(* CODESYS project Example15_PLC.project

Project tree, tasks and I/O mapping:
  Device : CODESYS Control Win V3, 3S - Smart Software Solutions GmbH, order no. 305021, version 3.5.7.0
    application Application
      libraries: Standard, * (System)
      task MainTask (cyclic, interval t#20ms, priority 1) calls PLC_PRG
      program PLC_PRG [ST]
      global variables GVL
      function block FB_G4LTL [ST]
    Ethernet : Ethernet, 3S - Smart Software Solutions GmbH, version 3.5.7.0
      Modbus_TCP_Master : Modbus TCP Master, 3S - Smart Software Solutions GmbH, version 3.5.6.0
          settings: AutoReconnect = TRUE
        Modbus_TCP_Slave : Modbus TCP Slave, 3S - Smart Software Solutions GmbH, version 3.5.7.0
            settings: Unit-ID = 1; IPAddress = [127, 0, 0, 1]; Channel 0.Function Code = 4; Channel 0.Read Offset = 16#0000; Channel 0.Read Length = 1; Channel 0.Write Offset = 0; Channel 0.Write Length = 0; Channel 0.Cycle Time = 100; Channel 1.Function Code = 4; Channel 1.Read Offset = 16#0001; Channel 1.Read Length = 1; Channel 1.Write Offset = 0; Channel 1.Write Length = 0; Channel 1.Cycle Time = 100; Channel 2.Function Code = 4; Channel 2.Read Offset = 16#0002; Channel 2.Read Length = 1; Channel 2.Write Offset = 0; Channel 2.Write Length = 0; Channel 2.Cycle Time = 100; Channel 3.Function Code = 4; Channel 3.Read Offset = 16#0003; Channel 3.Read Length = 1; Channel 3.Write Offset = 0; Channel 3.Write Length = 0; Channel 3.Cycle Time = 100; Channel 4.Function Code = 4; Channel 4.Read Offset = 16#0004; Channel 4.Read Length = 1; Channel 4.Write Offset = 0; Channel 4.Write Length = 0; Channel 4.Cycle Time = 100; Channel 5.Function Code = 6; Channel 5.Read Offset = 0; Channel 5.Read Length = 0; Channel 5.Write Offset = 16#0000; Channel 5.Write Length = 1; Channel 5.Cycle Time = 100; Channel 6.Function Code = 6; Channel 6.Read Offset = 0;
              Channel 6.Read Length = 0; Channel 6.Write Offset = 16#0002; Channel 6.Write Length = 1; Channel 6.Cycle Time = 100; Channel 7.Function Code = 6; Channel 7.Read Offset = 0; Channel 7.Read Length = 0; Channel 7.Write Offset = 16#0003; Channel 7.Write Length = 1; Channel 7.Cycle Time = 100; Channel 8.Function Code = 6; Channel 8.Read Offset = 0; Channel 8.Read Length = 0; Channel 8.Write Offset = 16#0004; Channel 8.Write Length = 1; Channel 8.Cycle Time = 100; Channel 9.Function Code = 6; Channel 9.Read Offset = 0; Channel 9.Read Length = 0; Channel 9.Write Offset = 16#0001; Channel 9.Write Length = 1; Channel 9.Cycle Time = 100; Channel 10.Function Code = 4; Channel 10.Read Offset = 16#0005; Channel 10.Read Length = 1; Channel 10.Write Offset = 0; Channel 10.Write Length = 0; Channel 10.Cycle Time = 100
            input  Application.dIn0 : BOOL  // Channel 0.Channel 0.Bit0
            input  Application.dIn1 : BOOL  // Channel 1.Channel 1.Bit0
            input  Application.dIn2 : BOOL  // Channel 2.Channel 2.Bit0
            input  Application.dIn3 : BOOL  // Channel 3.Channel 3.Bit0
            input  Application.dIn4 : BOOL  // Channel 4.Channel 4.Bit0
            output Application.dOut0 : BOOL  // Channel 5.Channel 5.Bit0
            output Application.dOut2 : BOOL  // Channel 6.Channel 6.Bit0
            output Application.dOut3 : BOOL  // Channel 7.Channel 7.Bit0
            output Application.dOut4 : BOOL  // Channel 8.Channel 8.Bit0
            output Application.dOut1 : BOOL  // Channel 9.Channel 9.Bit0
            input  Application.dIn5 : BOOL  // Channel 10.Channel 10.Bit0
            unmapped channels: Channel 0, Channel 1, Channel 2, Channel 3, Channel 4, Channel 5, Channel 6, Channel 7, Channel 8, Channel 9, Channel 10
*)

// Device/Application/GVL
VAR_GLOBAL
	
dIn0 : BOOL;
dIn1 : BOOL;
dIn2 : BOOL;
dIn3 : BOOL;
dIn4 : BOOL;
dIn5 : BOOL;

dOut0 : BOOL;
dOut1 : BOOL; 
dOut2 : BOOL; 
dOut3 : BOOL; 
dOut4 : BOOL; 
END_VAR

// Device/Application/PLC_PRG
PROGRAM PLC_PRG

VAR 
	fb: FB_G4LTL;
	
END_VAR


// Direct looping
// Assign pins (from global variable to function block) 
fb.x0 := dIn0;
fb.x1 := dIn1;
fb.x2 := dIn2;

// Assign pins (from function block to global variable)
dOut0 := fb.y0;
dOut1 := fb.y1;

// Run the function block
fb();

END_PROGRAM

// Device/Application/FB_G4LTL
FUNCTION_BLOCK FB_G4LTL
  (* Variable definition *)
   VAR_INPUT
      x0	: BOOL;
      x1	: BOOL;
      x2	: BOOL;
   END_VAR
   VAR_OUTPUT
      y0	: BOOL;
      y1	: BOOL;
   END_VAR
   VAR
   (* The total number of states equals to 100 *)
      cstate58	: LINT := 0;
      t0	: TON;
      t0_reset	: BOOL := FALSE;
      t0_up	: BOOL := FALSE;
      t0_start	: BOOL := FALSE;
	  
	  T0_VALUE	: TIME := TIME#7S;
   END_VAR

  (* Control logic *)
CASE cstate58 OF
1410:
    IF ((x0 = FALSE) AND  (x1 = FALSE) AND  (x2 = FALSE) AND  (t0.Q = FALSE)) THEN 
        cstate58 := 1220; y0 := FALSE; y1 := FALSE; t0_start := FALSE; 
    ELSIF ((x0 = FALSE) AND  (x1 = FALSE) AND  (x2 = FALSE) AND  (t0.Q = TRUE)) THEN 
        cstate58 := 1218; y0 := FALSE; y1 := FALSE; t0_start := FALSE; 
    ELSIF ((x0 = FALSE) AND  (x1 = FALSE) AND  (x2 = TRUE) AND  (t0.Q = FALSE)) THEN 
        cstate58 := 1412; y0 := FALSE; y1 := FALSE; t0_start := FALSE; 
    ELSIF ((x0 = FALSE) AND  (x1 = FALSE) AND  (x2 = TRUE) AND  (t0.Q = TRUE)) THEN 
        cstate58 := 1410; y0 := FALSE; y1 := FALSE; t0_start := FALSE; 
    ELSIF ((x0 = FALSE) AND  (x1 = TRUE) AND  (x2 = FALSE) AND  (t0.Q = FALSE)) THEN 
        cstate58 := 1220; y0 := FALSE; y1 := FALSE; t0_start := FALSE; 
    ELSIF ((x0 = FALSE) AND  (x1 = TRUE) AND  (x2 = FALSE) AND  (t0.Q = TRUE)) THEN 
        cstate58 := 1218; y0 := FALSE; y1 := FALSE; t0_start := FALSE; 
    ELSIF ((x0 = FALSE) AND  (x1 = TRUE) AND  (x2 = TRUE) AND  (t0.Q = FALSE)) THEN 
        cstate58 := 1412; y0 := FALSE; y1 := FALSE; t0_start := FALSE; 
    ELSIF ((x0 = FALSE) AND  (x1 = TRUE) AND  (x2 = TRUE) AND  (t0.Q = TRUE)) THEN 
        cstate58 := 1410; y0 := FALSE; y1 := FALSE; t0_start := FALSE; 
    ELSIF ((x0 = TRUE) AND  (x1 = FALSE) AND  (x2 = FALSE) AND  (t0.Q = FALSE)) THEN 
        cstate58 := 5192; y0 := TRUE; y1 := FALSE; t0_start := FALSE; 
    ELSIF ((x0 = TRUE) AND  (x1 = FALSE) AND  (x2 = FALSE) AND  (t0.Q = TRUE)) THEN 
        cstate58 := 5186; y0 := TRUE; y1 := FALSE; t0_start := FALSE; 
    ELSIF ((x0 = TRUE) AND  (x1 = FALSE) AND  (x2 = TRUE) AND  (t0.Q = FALSE)) THEN 
        cstate58 := 3848; y0 := FALSE; y1 := FALSE; t0_start := FALSE; 
    ELSIF ((x0 = TRUE) AND  (x1 = FALSE) AND  (x2 = TRUE) AND  (t0.Q = TRUE)) THEN 
        cstate58 := 3842; y0 := FALSE; y1 := FALSE; t0_start := FALSE; 
    ELSIF ((x0 = TRUE) AND  (x1 = TRUE) AND  (x2 = FALSE) AND  (t0.Q = FALSE)) THEN 
        cstate58 := 4678; y0 := TRUE; y1 := FALSE; t0_start := FALSE; 
    ELSIF ((x0 = TRUE) AND  (x1 = TRUE) AND  (x2 = FALSE) AND  (t0.Q = TRUE)) THEN 
        cstate58 := 4674; y0 := TRUE; y1 := FALSE; t0_start := FALSE; 
    ELSIF ((x0 = TRUE) AND  (x1 = TRUE) AND  (x2 = TRUE) AND  (t0.Q = FALSE)) THEN 
        cstate58 := 2502; y0 := FALSE; y1 := FALSE; t0_start := FALSE; 
    ELSIF ((x0 = TRUE) AND  (x1 = TRUE) AND  (x2 = TRUE) AND  (t0.Q = TRUE)) THEN 
        cstate58 := 2498; y0 := FALSE; y1 := FALSE; t0_start := FALSE; 
    END_IF;
6558:
    IF ((x0 = FALSE) AND  (x1 = FALSE) AND  (x2 = FALSE) AND  (t0.Q = FALSE)) THEN 
        cstate58 := 6366; y0 := FALSE; y1 := TRUE; t0_start := FALSE; 
    ELSIF ((x0 = FALSE) AND  (x1 = FALSE) AND  (x2 = FALSE) AND  (t0.Q = TRUE)) THEN 
        cstate58 := 6354; y0 := FALSE; y1 := TRUE; t0_start := FALSE; 
    ELSIF ((x0 = FALSE) AND  (x1 = FALSE) AND  (x2 = TRUE) AND  (t0.Q = FALSE)) THEN 
        cstate58 := 6558; y0 := FALSE; y1 := TRUE; t0_start := FALSE; 
    ELSIF ((x0 = FALSE) AND  (x1 = FALSE) AND  (x2 = TRUE) AND  (t0.Q = TRUE)) THEN 
        cstate58 := 6546; y0 := FALSE; y1 := TRUE; t0_start := FALSE; 
    ELSIF ((x0 = FALSE) AND  (x1 = TRUE) AND  (x2 = FALSE) AND  (t0.Q = FALSE)) THEN 
        cstate58 := 6340; y0 := FALSE; y1 := FALSE; t0_start := FALSE; 
    ELSIF ((x0 = FALSE) AND  (x1 = TRUE) AND  (x2 = FALSE) AND  (t0.Q = TRUE)) THEN 
        cstate58 := 6338; y0 := FALSE; y1 := FALSE; t0_start := FALSE; 
    ELSIF ((x0 = FALSE) AND  (x1 = TRUE) AND  (x2 = TRUE) AND  (t0.Q = FALSE)) THEN 
        cstate58 := 6532; y0 := FALSE; y1 := FALSE; t0_start := FALSE; 
    ELSIF ((x0 = FALSE) AND  (x1 = TRUE) AND  (x2 = TRUE) AND  (t0.Q = TRUE)) THEN 
        cstate58 := 6530; y0 := FALSE; y1 := FALSE; t0_start := FALSE; 
    ELSIF ((x0 = TRUE) AND  (x1 = FALSE) AND  (x2 = FALSE) AND  (t0.Q = FALSE)) THEN 
        cstate58 := 4168; y0 := TRUE; y1 := FALSE; t0_start := FALSE; 
    ELSIF ((x0 = TRUE) AND  (x1 = FALSE) AND  (x2 = FALSE) AND  (t0.Q = TRUE)) THEN 
        cstate58 := 4162; y0 := TRUE; y1 := FALSE; t0_start := FALSE; 
    ELSIF ((x0 = TRUE) AND  (x1 = FALSE) AND  (x2 = TRUE) AND  (t0.Q = FALSE)) THEN 
        cstate58 := 2824; y0 := FALSE; y1 := FALSE; t0_start := FALSE; 
    ELSIF ((x0 = TRUE) AND  (x1 = FALSE) AND  (x2 = TRUE) AND  (t0.Q = TRUE)) THEN 
        cstate58 := 2818; y0 := FALSE; y1 := FALSE; t0_start := FALSE; 
    ELSIF ((x0 = TRUE) AND  (x1 = TRUE) AND  (x2 = FALSE) AND  (t0.Q = FALSE)) THEN 
        cstate58 := 4678; y0 := TRUE; y1 := FALSE; t0_start := FALSE; 
    ELSIF ((x0 = TRUE) AND  (x1 = TRUE) AND  (x2 = FALSE) AND  (t0.Q = TRUE)) THEN 
        cstate58 := 4674; y0 := TRUE; y1 := FALSE; t0_start := FALSE; 
    ELSIF ((x0 = TRUE) AND  (x1 = TRUE) AND  (x2 = TRUE) AND  (t0.Q = FALSE)) THEN 
        cstate58 := 2502; y0 := FALSE; y1 := FALSE; t0_start := FALSE; 
    ELSIF ((x0 = TRUE) AND  (x1 = TRUE) AND  (x2 = TRUE) AND  (t0.Q = TRUE)) THEN 
        cstate58 := 2498; y0 := FALSE; y1 := FALSE; t0_start := FALSE; 
    END_IF;
1412:
    IF ((x0 = FALSE) AND  (x1 = FALSE) AND  (x2 = FALSE) AND  (t0.Q = FALSE)) THEN 
        cstate58 := 1220; y0 := FALSE; y1 := FALSE; t0_start := FALSE; 
    ELSIF ((x0 = FALSE) AND  (x1 = FALSE) AND  (x2 = FALSE) AND  (t0.Q = TRUE)) THEN 
        cstate58 := 1226; y0 := FALSE; y1 := TRUE; t0_start := FALSE; 
    ELSIF ((x0 = FALSE) AND  (x1 = FALSE) AND  (x2 = TRUE) AND  (t0.Q = FALSE)) THEN 
        cstate58 := 1412; y0 := FALSE; y1 := FALSE; t0_start := FALSE; 
    ELSIF ((x0 = FALSE) AND  (x1 = FALSE) AND  (x2 = TRUE) AND  (t0.Q = TRUE)) THEN 
        cstate58 := 1418; y0 := FALSE; y1 := TRUE; t0_start := FALSE; 
    ELSIF ((x0 = FALSE) AND  (x1 = TRUE) AND  (x2 = FALSE) AND  (t0.Q = FALSE)) THEN 
        cstate58 := 1220; y0 := FALSE; y1 := FALSE; t0_start := FALSE; 
    ELSIF ((x0 = FALSE) AND  (x1 = TRUE) AND  (x2 = FALSE) AND  (t0.Q = TRUE)) THEN 
        cstate58 := 1218; y0 := FALSE; y1 := FALSE; t0_start := FALSE; 
    ELSIF ((x0 = FALSE) AND  (x1 = TRUE) AND  (x2 = TRUE) AND  (t0.Q = FALSE)) THEN 
        cstate58 := 1412; y0 := FALSE; y1 := FALSE; t0_start := FALSE; 
    ELSIF ((x0 = FALSE) AND  (x1 = TRUE) AND  (x2 = TRUE) AND  (t0.Q = TRUE)) THEN 
        cstate58 := 1410; y0 := FALSE; y1 := FALSE; t0_start := FALSE; 
    ELSIF ((x0 = TRUE) AND  (x1 = FALSE) AND  (x2 = FALSE) AND  (t0.Q = FALSE)) THEN 
        cstate58 := 5192; y0 := TRUE; y1 := FALSE; t0_start := FALSE; 
    ELSIF ((x0 = TRUE) AND  (x1 = FALSE) AND  (x2 = FALSE) AND  (t0.Q = TRUE)) THEN 
        cstate58 := 5186; y0 := TRUE; y1 := FALSE; t0_start := FALSE; 
    ELSIF ((x0 = TRUE) AND  (x1 = FALSE) AND  (x2 = TRUE) AND  (t0.Q = FALSE)) THEN 
        cstate58 := 3848; y0 := FALSE; y1 := FALSE; t0_start := FALSE; 
    ELSIF ((x0 = TRUE) AND  (x1 = FALSE) AND  (x2 = TRUE) AND  (t0.Q = TRUE)) THEN 
        cstate58 := 3842; y0 := FALSE; y1 := FALSE; t0_start := FALSE; 
    ELSIF ((x0 = TRUE) AND  (x1 = TRUE) AND  (x2 = FALSE) AND  (t0.Q = FALSE)) THEN 
        cstate58 := 4678; y0 := TRUE; y1 := FALSE; t0_start := FALSE; 
    ELSIF ((x0 = TRUE) AND  (x1 = TRUE) AND  (x2 = FALSE) AND  (t0.Q = TRUE)) THEN 
        cstate58 := 4674; y0 := TRUE; y1 := FALSE; t0_start := FALSE; 
    ELSIF ((x0 = TRUE) AND  (x1 = TRUE) AND  (x2 = TRUE) AND  (t0.Q = FALSE)) THEN 
        cstate58 := 2502; y0 := FALSE; y1 := FALSE; t0_start := FALSE; 
    ELSIF ((x0 = TRUE) AND  (x1 = TRUE) AND  (x2 = TRUE) AND  (t0.Q = TRUE)) THEN 
        cstate58 := 2498; y0 := FALSE; y1 := FALSE; t0_start := FALSE; 
    END_IF;
1418:
    IF ((x0 = FALSE) AND  (x1 = FALSE) AND  (x2 = FALSE) AND  (t0.Q = FALSE)) THEN 
        cstate58 := 1238; y0 := FALSE; y1 := TRUE; t0_start := FALSE; 
    ELSIF ((x0 = FALSE) AND  (x1 = FALSE) AND  (x2 = FALSE) AND  (t0.Q = TRUE)) THEN 
        cstate58 := 1226; y0 := FALSE; y1 := TRUE; t0_start := FALSE; 
    ELSIF ((x0 = FALSE) AND  (x1 = FALSE) AND  (x2 = TRUE) AND  (t0.Q = FALSE)) THEN 
        cstate58 := 1430; y0 := FALSE; y1 := TRUE; t0_start := FALSE; 
    ELSIF ((x0 = FALSE) AND  (x1 = FALSE) AND  (x2 = TRUE) AND  (t0.Q = TRUE)) THEN 
        cstate58 := 1418; y0 := FALSE; y1 := TRUE; t0_start := FALSE; 
    ELSIF ((x0 = FALSE) AND  (x1 = TRUE) AND  (x2 = FALSE) AND  (t0.Q = FALSE)) THEN 
        cstate58 := 1220; y0 := FALSE; y1 := FALSE; t0_start := FALSE; 
    ELSIF ((x0 = FALSE) AND  (x1 = TRUE) AND  (x2 = FALSE) AND  (t0.Q = TRUE)) THEN 
        cstate58 := 1218; y0 := FALSE; y1 := FALSE; t0_start := FALSE; 
    ELSIF ((x0 = FALSE) AND  (x1 = TRUE) AND  (x2 = TRUE) AND  (t0.Q = FALSE)) THEN 
        cstate58 := 1412; y0 := FALSE; y1 := FALSE; t0_start := FALSE; 
    ELSIF ((x0 = FALSE) AND  (x1 = TRUE) AND  (x2 = TRUE) AND  (t0.Q = TRUE)) THEN 
        cstate58 := 1410; y0 := FALSE; y1 := FALSE; t0_start := FALSE; 
    ELSIF ((x0 = TRUE) AND  (x1 = FALSE) AND  (x2 = FALSE) AND  (t0.Q = FALSE)) THEN 
        cstate58 := 5192; y0 := TRUE; y1 := FALSE; t0_start := FALSE; 
    ELSIF ((x0 = TRUE) AND  (x1 = FALSE) AND  (x2 = FALSE) AND  (t0.Q = TRUE)) THEN 
        cstate58 := 5186; y0 := TRUE; y1 := FALSE; t0_start := FALSE; 
    ELSIF ((x0 = TRUE) AND  (x1 = FALSE) AND  (x2 = TRUE) AND  (t0.Q = FALSE)) THEN 
        cstate58 := 3848; y0 := FALSE; y1 := FALSE; t0_start := FALSE; 
    ELSIF ((x0 = TRUE) AND  (x1 = FALSE) AND  (x2 = TRUE) AND  (t0.Q = TRUE)) THEN 
        cstate58 := 3842; y0 := FALSE; y1 := FALSE; t0_start := FALSE; 
    ELSIF ((x0 = TRUE) AND  (x1 = TRUE) AND  (x2 = FALSE) AND  (t0.Q = FALSE)) THEN 
        cstate58 := 4678; y0 := TRUE; y1 := FALSE; t0_start := FALSE; 
    ELSIF ((x0 = TRUE) AND  (x1 = TRUE) AND  (x2 = FALSE) AND  (t0.Q = TRUE)) THEN 
        cstate58 := 4674; y0 := TRUE; y1 := FALSE; t0_start := FALSE; 
    ELSIF ((x0 = TRUE) AND  (x1 = TRUE) AND  (x2 = TRUE) AND  (t0.Q = FALSE)) THEN 
        cstate58 := 2502; y0 := FALSE; y1 := FALSE; t0_start := FALSE; 
    ELSIF ((x0 = TRUE) AND  (x1 = TRUE) AND  (x2 = TRUE) AND  (t0.Q = TRUE)) THEN 
        cstate58 := 2498; y0 := FALSE; y1 := FALSE; t0_start := FALSE; 
    END_IF;
7490:
    IF ((x0 = FALSE) AND  (x1 = FALSE) AND  (x2 = FALSE) AND  (t0.Q = FALSE)) THEN 
        cstate58 := 7428; y0 := FALSE; y1 := FALSE; t0_start := FALSE; 
    ELSIF ((x0 = FALSE) AND  (x1 = FALSE) AND  (x2 = FALSE) AND  (t0.Q = TRUE)) THEN 
        cstate58 := 7362; y0 := FALSE; y1 := FALSE; t0_start := FALSE; 
    ELSIF ((x0 = FALSE) AND  (x1 = FALSE) AND  (x2 = TRUE) AND  (t0.Q = FALSE)) THEN 
        cstate58 := 7492; y0 := FALSE; y1 := FALSE; t0_start := FALSE; 
    ELSIF ((x0 = FALSE) AND  (x1 = FALSE) AND  (x2 = TRUE) AND  (t0.Q = TRUE)) THEN 
        cstate58 := 7554; y0 := FALSE; y1 := FALSE; t0_start := FALSE; 
    ELSIF ((x0 = FALSE) AND  (x1 = TRUE) AND  (x2 = FALSE) AND  (t0.Q = FALSE)) THEN 
        cstate58 := 6404; y0 := FALSE; y1 := FALSE; t0_start := FALSE; 
    ELSIF ((x0 = FALSE) AND  (x1 = TRUE) AND  (x2 = FALSE) AND  (t0.Q = TRUE)) THEN 
        cstate58 := 6338; y0 := FALSE; y1 := FALSE; t0_start := FALSE; 
    ELSIF ((x0 = FALSE) AND  (x1 = TRUE) AND  (x2 = TRUE) AND  (t0.Q = FALSE)) THEN 
        cstate58 := 6468; y0 := FALSE; y1 := FALSE; t0_start := FALSE; 
    ELSIF ((x0 = FALSE) AND  (x1 = TRUE) AND  (x2 = TRUE) AND  (t0.Q = TRUE)) THEN 
        cstate58 := 6530; y0 := FALSE; y1 := FALSE; t0_start := FALSE; 
    ELSIF ((x0 = TRUE) AND  (x1 = FALSE) AND  (x2 = FALSE) AND  (t0.Q = FALSE)) THEN 
        cstate58 := 5256; y0 := TRUE; y1 := FALSE; t0_start := FALSE; 
    ELSIF ((x0 = TRUE) AND  (x1 = FALSE) AND  (x2 = FALSE) AND  (t0.Q = TRUE)) THEN 
        cstate58 := 5186; y0 := TRUE; y1 := FALSE; t0_start := FALSE; 
    ELSIF ((x0 = TRUE) AND  (x1 = FALSE) AND  (x2 = TRUE) AND  (t0.Q = FALSE)) THEN 
        cstate58 := 3784; y0 := FALSE; y1 := FALSE; t0_start := FALSE; 
    ELSIF ((x0 = TRUE) AND  (x1 = FALSE) AND  (x2 = TRUE) AND  (t0.Q = TRUE)) THEN 
        cstate58 := 3842; y0 := FALSE; y1 := FALSE; t0_start := FALSE; 
    ELSIF ((x0 = TRUE) AND  (x1 = TRUE) AND  (x2 = FALSE) AND  (t0.Q = FALSE)) THEN 
        cstate58 := 4742; y0 := TRUE; y1 := FALSE; t0_start := FALSE; 
    ELSIF ((x0 = TRUE) AND  (x1 = TRUE) AND  (x2 = FALSE) AND  (t0.Q = TRUE)) THEN 
        cstate58 := 4674; y0 := TRUE; y1 := FALSE; t0_start := FALSE; 
    ELSIF ((x0 = TRUE) AND  (x1 = TRUE) AND  (x2 = TRUE) AND  (t0.Q = FALSE)) THEN 
        cstate58 := 2566; y0 := FALSE; y1 := FALSE; t0_start := FALSE; 
    ELSIF ((x0 = TRUE) AND  (x1 = TRUE) AND  (x2 = TRUE) AND  (t0.Q = TRUE)) THEN 
        cstate58 := 2498; y0 := FALSE; y1 := FALSE; t0_start := FALSE; 
    END_IF;
7492:
    IF ((x0 = FALSE) AND  (x1 = FALSE) AND  (x2 = FALSE) AND  (t0.Q = FALSE)) THEN 
        cstate58 := 7428; y0 := FALSE; y1 := FALSE; t0_start := FALSE; 
    ELSIF ((x0 = FALSE) AND  (x1 = FALSE) AND  (x2 = FALSE) AND  (t0.Q = TRUE)) THEN 
        cstate58 := 7370; y0 := FALSE; y1 := TRUE; t0_start := FALSE; 
    ELSIF ((x0 = FALSE) AND  (x1 = FALSE) AND  (x2 = TRUE) AND  (t0.Q = FALSE)) THEN 
        cstate58 := 7492; y0 := FALSE; y1 := FALSE; t0_start := FALSE; 
    ELSIF ((x0 = FALSE) AND  (x1 = FALSE) AND  (x2 = TRUE) AND  (t0.Q = TRUE)) THEN 
        cstate58 := 7562; y0 := FALSE; y1 := TRUE; t0_start := FALSE; 
    ELSIF ((x0 = FALSE) AND  (x1 = TRUE) AND  (x2 = FALSE) AND  (t0.Q = FALSE)) THEN 
        cstate58 := 6404; y0 := FALSE; y1 := FALSE; t0_start := FALSE; 
    ELSIF ((x0 = FALSE) AND  (x1 = TRUE) AND  (x2 = FALSE) AND  (t0.Q = TRUE)) THEN 
        cstate58 := 6338; y0 := FALSE; y1 := FALSE; t0_start := FALSE; 
    ELSIF ((x0 = FALSE) AND  (x1 = TRUE) AND  (x2 = TRUE) AND  (t0.Q = FALSE)) THEN 
        cstate58 := 6468; y0 := FALSE; y1 := FALSE; t0_start := FALSE; 
    ELSIF ((x0 = FALSE) AND  (x1 = TRUE) AND  (x2 = TRUE) AND  (t0.Q = TRUE)) THEN 
        cstate58 := 6530; y0 := FALSE; y1 := FALSE; t0_start := FALSE; 
    ELSIF ((x0 = TRUE) AND  (x1 = FALSE) AND  (x2 = FALSE) AND  (t0.Q = FALSE)) THEN 
        cstate58 := 5256; y0 := TRUE; y1 := FALSE; t0_start := FALSE; 
    ELSIF ((x0 = TRUE) AND  (x1 = FALSE) AND  (x2 = FALSE) AND  (t0.Q = TRUE)) THEN 
        cstate58 := 5186; y0 := TRUE; y1 := FALSE; t0_start := FALSE; 
    ELSIF ((x0 = TRUE) AND  (x1 = FALSE) AND  (x2 = TRUE) AND  (t0.Q = FALSE)) THEN 
        cstate58 := 3784; y0 := FALSE; y1 := FALSE; t0_start := FALSE; 
    ELSIF ((x0 = TRUE) AND  (x1 = FALSE) AND  (x2 = TRUE) AND  (t0.Q = TRUE)) THEN 
        cstate58 := 3842; y0 := FALSE; y1 := FALSE; t0_start := FALSE; 
    ELSIF ((x0 = TRUE) AND  (x1 = TRUE) AND  (x2 = FALSE) AND  (t0.Q = FALSE)) THEN 
        cstate58 := 4742; y0 := TRUE; y1 := FALSE; t0_start := FALSE; 
    ELSIF ((x0 = TRUE) AND  (x1 = TRUE) AND  (x2 = FALSE) AND  (t0.Q = TRUE)) THEN 
        cstate58 := 4674; y0 := TRUE; y1 := FALSE; t0_start := FALSE; 
    ELSIF ((x0 = TRUE) AND  (x1 = TRUE) AND  (x2 = TRUE) AND  (t0.Q = FALSE)) THEN 
        cstate58 := 2566; y0 := FALSE; y1 := FALSE; t0_start := FALSE; 
    ELSIF ((x0 = TRUE) AND  (x1 = TRUE) AND  (x2 = TRUE) AND  (t0.Q = TRUE)) THEN 
        cstate58 := 2498; y0 := FALSE; y1 := FALSE; t0_start := FALSE; 
    END_IF;
6492:
    IF ((x0 = FALSE) AND  (x1 = FALSE) AND  (x2 = FALSE) AND  (t0.Q = FALSE)) THEN 
        cstate58 := 6428; y0 := FALSE; y1 := TRUE; t0_start := FALSE; 
    ELSIF ((x0 = FALSE) AND  (x1 = FALSE) AND  (x2 = FALSE) AND  (t0.Q = TRUE)) THEN 
        cstate58 := 6350; y0 := FALSE; y1 := TRUE; t0_start := FALSE; 
    ELSIF ((x0 = FALSE) AND  (x1 = FALSE) AND  (x2 = TRUE) AND  (t0.Q = FALSE)) THEN 
        cstate58 := 6492; y0 := FALSE; y1 := TRUE; t0_start := FALSE; 
    ELSIF ((x0 = FALSE) AND  (x1 = FALSE) AND  (x2 = TRUE) AND  (t0.Q = TRUE)) THEN 
        cstate58 := 6542; y0 := FALSE; y1 := TRUE; t0_start := FALSE; 
    ELSIF ((x0 = FALSE) AND  (x1 = TRUE) AND  (x2 = FALSE) AND  (t0.Q = FALSE)) THEN 
        cstate58 := 6404; y0 := FALSE; y1 := FALSE; t0_start := FALSE; 
    ELSIF ((x0 = FALSE) AND  (x1 = TRUE) AND  (x2 = FALSE) AND  (t0.Q = TRUE)) THEN 
        cstate58 := 6338; y0 := FALSE; y1 := FALSE; t0_start := FALSE; 
    ELSIF ((x0 = FALSE) AND  (x1 = TRUE) AND  (x2 = TRUE) AND  (t0.Q = FALSE)) THEN 
        cstate58 := 6468; y0 := FALSE; y1 := FALSE; t0_start := FALSE; 
    ELSIF ((x0 = FALSE) AND  (x1 = TRUE) AND  (x2 = TRUE) AND  (t0.Q = TRUE)) THEN 
        cstate58 := 6530; y0 := FALSE; y1 := FALSE; t0_start := FALSE; 
    ELSIF ((x0 = TRUE) AND  (x1 = FALSE) AND  (x2 = FALSE) AND  (t0.Q = FALSE)) THEN 
        cstate58 := 4232; y0 := TRUE; y1 := FALSE; t0_start := FALSE; 
    ELSIF ((x0 = TRUE) AND  (x1 = FALSE) AND  (x2 = FALSE) AND  (t0.Q = TRUE)) THEN 
        cstate58 := 4162; y0 := TRUE; y1 := FALSE; t0_start := FALSE; 
    ELSIF ((x0 = TRUE) AND  (x1 = FALSE) AND  (x2 = TRUE) AND  (t0.Q = FALSE)) THEN 
        cstate58 := 2760; y0 := FALSE; y1 := FALSE; t0_start := FALSE; 
    ELSIF ((x0 = TRUE) AND  (x1 = FALSE) AND  (x2 = TRUE) AND  (t0.Q = TRUE)) THEN 
        cstate58 := 2818; y0 := FALSE; y1 := FALSE; t0_start := FALSE; 
    ELSIF ((x0 = TRUE) AND  (x1 = TRUE) AND  (x2 = FALSE) AND  (t0.Q = FALSE)) THEN 
        cstate58 := 4742; y0 := TRUE; y1 := FALSE; t0_start := FALSE; 
    ELSIF ((x0 = TRUE) AND  (x1 = TRUE) AND  (x2 = FALSE) AND  (t0.Q = TRUE)) THEN 
        cstate58 := 4674; y0 := TRUE; y1 := FALSE; t0_start := FALSE; 
    ELSIF ((x0 = TRUE) AND  (x1 = TRUE) AND  (x2 = TRUE) AND  (t0.Q = FALSE)) THEN 
        cstate58 := 2566; y0 := FALSE; y1 := FALSE; t0_start := FALSE; 
    ELSIF ((x0 = TRUE) AND  (x1 = TRUE) AND  (x2 = TRUE) AND  (t0.Q = TRUE)) THEN 
        cstate58 := 2498; y0 := FALSE; y1 := FALSE; t0_start := FALSE; 
    END_IF;
6350:
    IF ((x0 = FALSE) AND  (x1 = FALSE) AND  (x2 = FALSE) AND  (t0.Q = FALSE)) THEN 
        cstate58 := 6362; y0 := FALSE; y1 := TRUE; t0_start := FALSE; 
    ELSIF ((x0 = FALSE) AND  (x1 = FALSE) AND  (x2 = FALSE) AND  (t0.Q = TRUE)) THEN 
        cstate58 := 6350; y0 := FALSE; y1 := TRUE; t0_start := FALSE; 
    ELSIF ((x0 = FALSE) AND  (x1 = FALSE) AND  (x2 = TRUE) AND  (t0.Q = FALSE)) THEN 
        cstate58 := 6492; y0 := FALSE; y1 := TRUE; t0_start := TRUE; t0_up := FALSE; 
    ELSIF ((x0 = FALSE) AND  (x1 = FALSE) AND  (x2 = TRUE) AND  (t0.Q = TRUE)) THEN 
        cstate58 := 6480; y0 := FALSE; y1 := TRUE; t0_start := TRUE; t0_up := FALSE; 
    ELSIF ((x0 = FALSE) AND  (x1 = TRUE) AND  (x2 = FALSE) AND  (t0.Q = FALSE)) THEN 
        cstate58 := 6340; y0 := FALSE; y1 := FALSE; t0_start := FALSE; 
    ELSIF ((x0 = FALSE) AND  (x1 = TRUE) AND  (x2 = FALSE) AND  (t0.Q = TRUE)) THEN 
        cstate58 := 6338; y0 := FALSE; y1 := FALSE; t0_start := FALSE; 
    ELSIF ((x0 = FALSE) AND  (x1 = TRUE) AND  (x2 = TRUE) AND  (t0.Q = FALSE)) THEN 
        cstate58 := 6468; y0 := FALSE; y1 := FALSE; t0_start := TRUE; t0_up := FALSE; 
    ELSIF ((x0 = FALSE) AND  (x1 = TRUE) AND  (x2 = TRUE) AND  (t0.Q = TRUE)) THEN 
        cstate58 := 6466; y0 := FALSE; y1 := FALSE; t0_start := TRUE; t0_up := FALSE; 
    ELSIF ((x0 = TRUE) AND  (x1 = FALSE) AND  (x2 = FALSE) AND  (t0.Q = FALSE)) THEN 
        cstate58 := 4168; y0 := TRUE; y1 := FALSE; t0_start := FALSE; 
    ELSIF ((x0 = TRUE) AND  (x1 = FALSE) AND  (x2 = FALSE) AND  (t0.Q = TRUE)) THEN 
        cstate58 := 4162; y0 := TRUE; y1 := FALSE; t0_start := FALSE; 
    ELSIF ((x0 = TRUE) AND  (x1 = FALSE) AND  (x2 = TRUE) AND  (t0.Q = FALSE)) THEN 
        cstate58 := 2760; y0 := FALSE; y1 := FALSE; t0_start := TRUE; t0_up := FALSE; 
    ELSIF ((x0 = TRUE) AND  (x1 = FALSE) AND  (x2 = TRUE) AND  (t0.Q = TRUE)) THEN 
        cstate58 := 2754; y0 := FALSE; y1 := FALSE; t0_start := TRUE; t0_up := FALSE; 
    ELSIF ((x0 = TRUE) AND  (x1 = TRUE) AND  (x2 = FALSE) AND  (t0.Q = FALSE)) THEN 
        cstate58 := 4678; y0 := TRUE; y1 := FALSE; t0_start := FALSE; 
    ELSIF ((x0 = TRUE) AND  (x1 = TRUE) AND  (x2 = FALSE) AND  (t0.Q = TRUE)) THEN 
        cstate58 := 4674; y0 := TRUE; y1 := FALSE; t0_start := FALSE; 
    ELSIF ((x0 = TRUE) AND  (x1 = TRUE) AND  (x2 = TRUE) AND  (t0.Q = FALSE)) THEN 
        cstate58 := 2566; y0 := FALSE; y1 := FALSE; t0_start := TRUE; t0_up := FALSE; 
    ELSIF ((x0 = TRUE) AND  (x1 = TRUE) AND  (x2 = TRUE) AND  (t0.Q = TRUE)) THEN 
        cstate58 := 2562; y0 := FALSE; y1 := FALSE; t0_start := TRUE; t0_up := FALSE; 
    END_IF;
6354:
    IF ((x0 = FALSE) AND  (x1 = FALSE) AND  (x2 = FALSE) AND  (t0.Q = FALSE)) THEN 
        cstate58 := 6366; y0 := FALSE; y1 := TRUE; t0_start := FALSE; 
    ELSIF ((x0 = FALSE) AND  (x1 = FALSE) AND  (x2 = FALSE) AND  (t0.Q = TRUE)) THEN 
        cstate58 := 6354; y0 := FALSE; y1 := TRUE; t0_start := FALSE; 
    ELSIF ((x0 = FALSE) AND  (x1 = FALSE) AND  (x2 = TRUE) AND  (t0.Q = FALSE)) THEN 
        cstate58 := 6496; y0 := FALSE; y1 := TRUE; t0_start := TRUE; t0_up := FALSE; 
    ELSIF ((x0 = FALSE) AND  (x1 = FALSE) AND  (x2 = TRUE) AND  (t0.Q = TRUE)) THEN 
        cstate58 := 6484; y0 := FALSE; y1 := TRUE; t0_start := TRUE; t0_up := FALSE; 
    ELSIF ((x0 = FALSE) AND  (x1 = TRUE) AND  (x2 = FALSE) AND  (t0.Q = FALSE)) THEN 
        cstate58 := 6340; y0 := FALSE; y1 := FALSE; t0_start := FALSE; 
    ELSIF ((x0 = FALSE) AND  (x1 = TRUE) AND  (x2 = FALSE) AND  (t0.Q = TRUE)) THEN 
        cstate58 := 6338; y0 := FALSE; y1 := FALSE; t0_start := FALSE; 
    ELSIF ((x0 = FALSE) AND  (x1 = TRUE) AND  (x2 = TRUE) AND  (t0.Q = FALSE)) THEN 
        cstate58 := 6468; y0 := FALSE; y1 := FALSE; t0_start := TRUE; t0_up := FALSE; 
    ELSIF ((x0 = FALSE) AND  (x1 = TRUE) AND  (x2 = TRUE) AND  (t0.Q = TRUE)) THEN 
        cstate58 := 6466; y0 := FALSE; y1 := FALSE; t0_start := TRUE; t0_up := FALSE; 
    ELSIF ((x0 = TRUE) AND  (x1 = FALSE) AND  (x2 = FALSE) AND  (t0.Q = FALSE)) THEN 
        cstate58 := 4168; y0 := TRUE; y1 := FALSE; t0_start := FALSE; 
    ELSIF ((x0 = TRUE) AND  (x1 = FALSE) AND  (x2 = FALSE) AND  (t0.Q = TRUE)) THEN 
        cstate58 := 4162; y0 := TRUE; y1 := FALSE; t0_start := FALSE; 
    ELSIF ((x0 = TRUE) AND  (x1 = FALSE) AND  (x2 = TRUE) AND  (t0.Q = FALSE)) THEN 
        cstate58 := 2760; y0 := FALSE; y1 := FALSE; t0_start := TRUE; t0_up := FALSE; 
    ELSIF ((x0 = TRUE) AND  (x1 = FALSE) AND  (x2 = TRUE) AND  (t0.Q = TRUE)) THEN 
        cstate58 := 2754; y0 := FALSE; y1 := FALSE; t0_start := TRUE; t0_up := FALSE; 
    ELSIF ((x0 = TRUE) AND  (x1 = TRUE) AND  (x2 = FALSE) AND  (t0.Q = FALSE)) THEN 
        cstate58 := 4678; y0 := TRUE; y1 := FALSE; t0_start := FALSE; 
    ELSIF ((x0 = TRUE) AND  (x1 = TRUE) AND  (x2 = FALSE) AND  (t0.Q = TRUE)) THEN 
        cstate58 := 4674; y0 := TRUE; y1 := FALSE; t0_start := FALSE; 
    ELSIF ((x0 = TRUE) AND  (x1 = TRUE) AND  (x2 = TRUE) AND  (t0.Q = FALSE)) THEN 
        cstate58 := 2566; y0 := FALSE; y1 := FALSE; t0_start := TRUE; t0_up := FALSE; 
    ELSIF ((x0 = TRUE) AND  (x1 = TRUE) AND  (x2 = TRUE) AND  (t0.Q = TRUE)) THEN 
        cstate58 := 2562; y0 := FALSE; y1 := FALSE; t0_start := TRUE; t0_up := FALSE; 
    END_IF;
6496:
    IF ((x0 = FALSE) AND  (x1 = FALSE) AND  (x2 = FALSE) AND  (t0.Q = FALSE)) THEN 
        cstate58 := 6432; y0 := FALSE; y1 := TRUE; t0_start := FALSE; 
    ELSIF ((x0 = FALSE) AND  (x1 = FALSE) AND  (x2 = FALSE) AND  (t0.Q = TRUE)) THEN 
        cstate58 := 6354; y0 := FALSE; y1 := TRUE; t0_start := FALSE; 
    ELSIF ((x0 = FALSE) AND  (x1 = FALSE) AND  (x2 = TRUE) AND  (t0.Q = FALSE)) THEN 
        cstate58 := 6496; y0 := FALSE; y1 := TRUE; t0_start := FALSE; 
    ELSIF ((x0 = FALSE) AND  (x1 = FALSE) AND  (x2 = TRUE) AND  (t0.Q = TRUE)) THEN 
        cstate58 := 6546; y0 := FALSE; y1 := TRUE; t0_start := FALSE; 
    ELSIF ((x0 = FALSE) AND  (x1 = TRUE) AND  (x2 = FALSE) AND  (t0.Q = FALSE)) THEN 
        cstate58 := 6404; y0 := FALSE; y1 := FALSE; t0_start := FALSE; 
    ELSIF ((x0 = FALSE) AND  (x1 = TRUE) AND  (x2 = FALSE) AND  (t0.Q = TRUE)) THEN 
        cstate58 := 6338; y0 := FALSE; y1 := FALSE; t0_start := FALSE; 
    ELSIF ((x0 = FALSE) AND  (x1 = TRUE) AND  (x2 = TRUE) AND  (t0.Q = FALSE)) THEN 
        cstate58 := 6468; y0 := FALSE; y1 := FALSE; t0_start := FALSE; 
    ELSIF ((x0 = FALSE) AND  (x1 = TRUE) AND  (x2 = TRUE) AND  (t0.Q = TRUE)) THEN 
        cstate58 := 6530; y0 := FALSE; y1 := FALSE; t0_start := FALSE; 
    ELSIF ((x0 = TRUE) AND  (x1 = FALSE) AND  (x2 = FALSE) AND  (t0.Q = FALSE)) THEN 
        cstate58 := 4232; y0 := TRUE; y1 := FALSE; t0_start := FALSE; 
    ELSIF ((x0 = TRUE) AND  (x1 = FALSE) AND  (x2 = FALSE) AND  (t0.Q = TRUE)) THEN 
        cstate58 := 4162; y0 := TRUE; y1 := FALSE; t0_start := FALSE; 
    ELSIF ((x0 = TRUE) AND  (x1 = FALSE) AND  (x2 = TRUE) AND  (t0.Q = FALSE)) THEN 
        cstate58 := 2760; y0 := FALSE; y1 := FALSE; t0_start := FALSE; 
    ELSIF ((x0 = TRUE) AND  (x1 = FALSE) AND  (x2 = TRUE) AND  (t0.Q = TRUE)) THEN 
        cstate58 := 2818; y0 := FALSE; y1 := FALSE; t0_start := FALSE; 
    ELSIF ((x0 = TRUE) AND  (x1 = TRUE) AND  (x2 = FALSE) AND  (t0.Q = FALSE)) THEN 
        cstate58 := 4742; y0 := TRUE; y1 := FALSE; t0_start := FALSE; 
    ELSIF ((x0 = TRUE) AND  (x1 = TRUE) AND  (x2 = FALSE) AND  (t0.Q = TRUE)) THEN 
        cstate58 := 4674; y0 := TRUE; y1 := FALSE; t0_start := FALSE; 
    ELSIF ((x0 = TRUE) AND  (x1 = TRUE) AND  (x2 = TRUE) AND  (t0.Q = FALSE)) THEN 
        cstate58 := 2566; y0 := FALSE; y1 := FALSE; t0_start := FALSE; 
    ELSIF ((x0 = TRUE) AND  (x1 = TRUE) AND  (x2 = TRUE) AND  (t0.Q = TRUE)) THEN 
        cstate58 := 2498; y0 := FALSE; y1 := FALSE; t0_start := FALSE; 
    END_IF;
6546:
    IF ((x0 = FALSE) AND  (x1 = FALSE) AND  (x2 = FALSE) AND  (t0.Q = FALSE)) THEN 
        cstate58 := 6366; y0 := FALSE; y1 := TRUE; t0_start := FALSE; 
    ELSIF ((x0 = FALSE) AND  (x1 = FALSE) AND  (x2 = FALSE) AND  (t0.Q = TRUE)) THEN 
        cstate58 := 6354; y0 := FALSE; y1 := TRUE; t0_start := FALSE; 
    ELSIF ((x0 = FALSE) AND  (x1 = FALSE) AND  (x2 = TRUE) AND  (t0.Q = FALSE)) THEN 
        cstate58 := 6558; y0 := FALSE; y1 := TRUE; t0_start := FALSE; 
    ELSIF ((x0 = FALSE) AND  (x1 = FALSE) AND  (x2 = TRUE) AND  (t0.Q = TRUE)) THEN 
        cstate58 := 6546; y0 := FALSE; y1 := TRUE; t0_start := FALSE; 
    ELSIF ((x0 = FALSE) AND  (x1 = TRUE) AND  (x2 = FALSE) AND  (t0.Q = FALSE)) THEN 
        cstate58 := 6340; y0 := FALSE; y1 := FALSE; t0_start := FALSE; 
    ELSIF ((x0 = FALSE) AND  (x1 = TRUE) AND  (x2 = FALSE) AND  (t0.Q = TRUE)) THEN 
        cstate58 := 6338; y0 := FALSE; y1 := FALSE; t0_start := FALSE; 
    ELSIF ((x0 = FALSE) AND  (x1 = TRUE) AND  (x2 = TRUE) AND  (t0.Q = FALSE)) THEN 
        cstate58 := 6532; y0 := FALSE; y1 := FALSE; t0_start := FALSE; 
    ELSIF ((x0 = FALSE) AND  (x1 = TRUE) AND  (x2 = TRUE) AND  (t0.Q = TRUE)) THEN 
        cstate58 := 6530; y0 := FALSE; y1 := FALSE; t0_start := FALSE; 
    ELSIF ((x0 = TRUE) AND  (x1 = FALSE) AND  (x2 = FALSE) AND  (t0.Q = FALSE)) THEN 
        cstate58 := 4168; y0 := TRUE; y1 := FALSE; t0_start := FALSE; 
    ELSIF ((x0 = TRUE) AND  (x1 = FALSE) AND  (x2 = FALSE) AND  (t0.Q = TRUE)) THEN 
        cstate58 := 4162; y0 := TRUE; y1 := FALSE; t0_start := FALSE; 
    ELSIF ((x0 = TRUE) AND  (x1 = FALSE) AND  (x2 = TRUE) AND  (t0.Q = FALSE)) THEN 
        cstate58 := 2824; y0 := FALSE; y1 := FALSE; t0_start := FALSE; 
    ELSIF ((x0 = TRUE) AND  (x1 = FALSE) AND  (x2 = TRUE) AND  (t0.Q = TRUE)) THEN 
        cstate58 := 2818; y0 := FALSE; y1 := FALSE; t0_start := FALSE; 
    ELSIF ((x0 = TRUE) AND  (x1 = TRUE) AND  (x2 = FALSE) AND  (t0.Q = FALSE)) THEN 
        cstate58 := 4678; y0 := TRUE; y1 := FALSE; t0_start := FALSE; 
    ELSIF ((x0 = TRUE) AND  (x1 = TRUE) AND  (x2 = FALSE) AND  (t0.Q = TRUE)) THEN 
        cstate58 := 4674; y0 := TRUE; y1 := FALSE; t0_start := FALSE; 
    ELSIF ((x0 = TRUE) AND  (x1 = TRUE) AND  (x2 = TRUE) AND  (t0.Q = FALSE)) THEN 
        cstate58 := 2502; y0 := FALSE; y1 := FALSE; t0_start := FALSE; 
    ELSIF ((x0 = TRUE) AND  (x1 = TRUE) AND  (x2 = TRUE) AND  (t0.Q = TRUE)) THEN 
        cstate58 := 2498; y0 := FALSE; y1 := FALSE; t0_start := FALSE; 
    END_IF;
1284:
    IF ((x0 = FALSE) AND  (x1 = FALSE) AND  (x2 = FALSE) AND  (t0.Q = FALSE)) THEN 
        cstate58 := 1284; y0 := FALSE; y1 := FALSE; t0_start := FALSE; 
    ELSIF ((x0 = FALSE) AND  (x1 = FALSE) AND  (x2 = FALSE) AND  (t0.Q = TRUE)) THEN 
        cstate58 := 1226; y0 := FALSE; y1 := TRUE; t0_start := FALSE; 
    ELSIF ((x0 = FALSE) AND  (x1 = FALSE) AND  (x2 = TRUE) AND  (t0.Q = FALSE)) THEN 
        cstate58 := 1348; y0 := FALSE; y1 := FALSE; t0_start := TRUE; t0_up := FALSE; 
    ELSIF ((x0 = FALSE) AND  (x1 = FALSE) AND  (x2 = TRUE) AND  (t0.Q = TRUE)) THEN 
        cstate58 := 1356; y0 := FALSE; y1 := TRUE; t0_start := TRUE; t0_up := FALSE; 
    ELSIF ((x0 = FALSE) AND  (x1 = TRUE) AND  (x2 = FALSE) AND  (t0.Q = FALSE)) THEN 
        cstate58 := 1284; y0 := FALSE; y1 := FALSE; t0_start := FALSE; 
    ELSIF ((x0 = FALSE) AND  (x1 = TRUE) AND  (x2 = FALSE) AND  (t0.Q = TRUE)) THEN 
        cstate58 := 1218; y0 := FALSE; y1 := FALSE; t0_start := FALSE; 
    ELSIF ((x0 = FALSE) AND  (x1 = TRUE) AND  (x2 = TRUE) AND  (t0.Q = FALSE)) THEN 
        cstate58 := 1348; y0 := FALSE; y1 := FALSE; t0_start := TRUE; t0_up := FALSE; 
    ELSIF ((x0 = FALSE) AND  (x1 = TRUE) AND  (x2 = TRUE) AND  (t0.Q = TRUE)) THEN 
        cstate58 := 1346; y0 := FALSE; y1 := FALSE; t0_start := TRUE; t0_up := FALSE; 
    ELSIF ((x0 = TRUE) AND  (x1 = FALSE) AND  (x2 = FALSE) AND  (t0.Q = FALSE)) THEN 
        cstate58 := 5256; y0 := TRUE; y1 := FALSE; t0_start := FALSE; 
    ELSIF ((x0 = TRUE) AND  (x1 = FALSE) AND  (x2 = FALSE) AND  (t0.Q = TRUE)) THEN 
        cstate58 := 5186; y0 := TRUE; y1 := FALSE; t0_start := FALSE; 
    ELSIF ((x0 = TRUE) AND  (x1 = FALSE) AND  (x2 = TRUE) AND  (t0.Q = FALSE)) THEN 
        cstate58 := 3784; y0 := FALSE; y1 := FALSE; t0_start := TRUE; t0_up := FALSE; 
    ELSIF ((x0 = TRUE) AND  (x1 = FALSE) AND  (x2 = TRUE) AND  (t0.Q = TRUE)) THEN 
        cstate58 := 3778; y0 := FALSE; y1 := FALSE; t0_start := TRUE; t0_up := FALSE; 
    ELSIF ((x0 = TRUE) AND  (x1 = TRUE) AND  (x2 = FALSE) AND  (t0.Q = FALSE)) THEN 
        cstate58 := 4742; y0 := TRUE; y1 := FALSE; t0_start := FALSE; 
    ELSIF ((x0 = TRUE) AND  (x1 = TRUE) AND  (x2 = FALSE) AND  (t0.Q = TRUE)) THEN 
        cstate58 := 4674; y0 := TRUE; y1 := FALSE; t0_start := FALSE; 
    ELSIF ((x0 = TRUE) AND  (x1 = TRUE) AND  (x2 = TRUE) AND  (t0.Q = FALSE)) THEN 
        cstate58 := 2566; y0 := FALSE; y1 := FALSE; t0_start := TRUE; t0_up := FALSE; 
    ELSIF ((x0 = TRUE) AND  (x1 = TRUE) AND  (x2 = TRUE) AND  (t0.Q = TRUE)) THEN 
        cstate58 := 2562; y0 := FALSE; y1 := FALSE; t0_start := TRUE; t0_up := FALSE; 
    END_IF;
3208:
    IF ((x0 = FALSE) AND  (x1 = FALSE) AND  (x2 = FALSE) AND  (t0.Q = FALSE)) THEN 
        cstate58 := 7428; y0 := FALSE; y1 := FALSE; t0_start := FALSE; 
    ELSIF ((x0 = FALSE) AND  (x1 = FALSE) AND  (x2 = FALSE) AND  (t0.Q = TRUE)) THEN 
        cstate58 := 7378; y0 := FALSE; y1 := TRUE; t0_start := FALSE; 
    ELSIF ((x0 = FALSE) AND  (x1 = FALSE) AND  (x2 = TRUE) AND  (t0.Q = FALSE)) THEN 
        cstate58 := 7492; y0 := FALSE; y1 := FALSE; t0_start := TRUE; t0_up := FALSE; 
    ELSIF ((x0 = FALSE) AND  (x1 = FALSE) AND  (x2 = TRUE) AND  (t0.Q = TRUE)) THEN 
        cstate58 := 7508; y0 := FALSE; y1 := TRUE; t0_start := TRUE; t0_up := FALSE; 
    ELSIF ((x0 = FALSE) AND  (x1 = TRUE) AND  (x2 = FALSE) AND  (t0.Q = FALSE)) THEN 
        cstate58 := 6404; y0 := FALSE; y1 := FALSE; t0_start := FALSE; 
    ELSIF ((x0 = FALSE) AND  (x1 = TRUE) AND  (x2 = FALSE) AND  (t0.Q = TRUE)) THEN 
        cstate58 := 6338; y0 := FALSE; y1 := FALSE; t0_start := FALSE; 
    ELSIF ((x0 = FALSE) AND  (x1 = TRUE) AND  (x2 = TRUE) AND  (t0.Q = FALSE)) THEN 
        cstate58 := 6468; y0 := FALSE; y1 := FALSE; t0_start := TRUE; t0_up := FALSE; 
    ELSIF ((x0 = FALSE) AND  (x1 = TRUE) AND  (x2 = TRUE) AND  (t0.Q = TRUE)) THEN 
        cstate58 := 6466; y0 := FALSE; y1 := FALSE; t0_start := TRUE; t0_up := FALSE; 
    ELSIF ((x0 = TRUE) AND  (x1 = FALSE) AND  (x2 = FALSE) AND  (t0.Q = FALSE)) THEN 
        cstate58 := 3208; y0 := FALSE; y1 := FALSE; t0_start := FALSE; 
    ELSIF ((x0 = TRUE) AND  (x1 = FALSE) AND  (x2 = FALSE) AND  (t0.Q = TRUE)) THEN 
        cstate58 := 3138; y0 := FALSE; y1 := FALSE; t0_start := FALSE; 
    ELSIF ((x0 = TRUE) AND  (x1 = FALSE) AND  (x2 = TRUE) AND  (t0.Q = FALSE)) THEN 
        cstate58 := 3784; y0 := FALSE; y1 := FALSE; t0_start := TRUE; t0_up := FALSE; 
    ELSIF ((x0 = TRUE) AND  (x1 = FALSE) AND  (x2 = TRUE) AND  (t0.Q = TRUE)) THEN 
        cstate58 := 3778; y0 := FALSE; y1 := FALSE; t0_start := TRUE; t0_up := FALSE; 
    ELSIF ((x0 = TRUE) AND  (x1 = TRUE) AND  (x2 = FALSE) AND  (t0.Q = FALSE)) THEN 
        cstate58 := 2694; y0 := FALSE; y1 := FALSE; t0_start := FALSE; 
    ELSIF ((x0 = TRUE) AND  (x1 = TRUE) AND  (x2 = FALSE) AND  (t0.Q = TRUE)) THEN 
        cstate58 := 2626; y0 := FALSE; y1 := FALSE; t0_start := FALSE; 
    ELSIF ((x0 = TRUE) AND  (x1 = TRUE) AND  (x2 = TRUE) AND  (t0.Q = FALSE)) THEN 
        cstate58 := 2566; y0 := FALSE; y1 := FALSE; t0_start := TRUE; t0_up := FALSE; 
    ELSIF ((x0 = TRUE) AND  (x1 = TRUE) AND  (x2 = TRUE) AND  (t0.Q = TRUE)) THEN 
        cstate58 := 2562; y0 := FALSE; y1 := FALSE; t0_start := TRUE; t0_up := FALSE; 
    END_IF;
3138:
    IF ((x0 = FALSE) AND  (x1 = FALSE) AND  (x2 = FALSE) AND  (t0.Q = FALSE)) THEN 
        cstate58 := 7364; y0 := FALSE; y1 := FALSE; t0_start := FALSE; 
    ELSIF ((x0 = FALSE) AND  (x1 = FALSE) AND  (x2 = FALSE) AND  (t0.Q = TRUE)) THEN 
        cstate58 := 7362; y0 := FALSE; y1 := FALSE; t0_start := FALSE; 
    ELSIF ((x0 = FALSE) AND  (x1 = FALSE) AND  (x2 = TRUE) AND  (t0.Q = FALSE)) THEN 
        cstate58 := 7492; y0 := FALSE; y1 := FALSE; t0_start := TRUE; t0_up := FALSE; 
    ELSIF ((x0 = FALSE) AND  (x1 = FALSE) AND  (x2 = TRUE) AND  (t0.Q = TRUE)) THEN 
        cstate58 := 7490; y0 := FALSE; y1 := FALSE; t0_start := TRUE; t0_up := FALSE; 
    ELSIF ((x0 = FALSE) AND  (x1 = TRUE) AND  (x2 = FALSE) AND  (t0.Q = FALSE)) THEN 
        cstate58 := 6340; y0 := FALSE; y1 := FALSE; t0_start := FALSE; 
    ELSIF ((x0 = FALSE) AND  (x1 = TRUE) AND  (x2 = FALSE) AND  (t0.Q = TRUE)) THEN 
        cstate58 := 6338; y0 := FALSE; y1 := FALSE; t0_start := FALSE; 
    ELSIF ((x0 = FALSE) AND  (x1 = TRUE) AND  (x2 = TRUE) AND  (t0.Q = FALSE)) THEN 
        cstate58 := 6468; y0 := FALSE; y1 := FALSE; t0_start := TRUE; t0_up := FALSE; 
    ELSIF ((x0 = FALSE) AND  (x1 = TRUE) AND  (x2 = TRUE) AND  (t0.Q = TRUE)) THEN 
        cstate58 := 6466; y0 := FALSE; y1 := FALSE; t0_start := TRUE; t0_up := FALSE; 
    ELSIF ((x0 = TRUE) AND  (x1 = FALSE) AND  (x2 = FALSE) AND  (t0.Q = FALSE)) THEN 
        cstate58 := 3144; y0 := FALSE; y1 := FALSE; t0_start := FALSE; 
    ELSIF ((x0 = TRUE) AND  (x1 = FALSE) AND  (x2 = FALSE) AND  (t0.Q = TRUE)) THEN 
        cstate58 := 3138; y0 := FALSE; y1 := FALSE; t0_start := FALSE; 
    ELSIF ((x0 = TRUE) AND  (x1 = FALSE) AND  (x2 = TRUE) AND  (t0.Q = FALSE)) THEN 
        cstate58 := 3784; y0 := FALSE; y1 := FALSE; t0_start := TRUE; t0_up := FALSE; 
    ELSIF ((x0 = TRUE) AND  (x1 = FALSE) AND  (x2 = TRUE) AND  (t0.Q = TRUE)) THEN 
        cstate58 := 3778; y0 := FALSE; y1 := FALSE; t0_start := TRUE; t0_up := FALSE; 
    ELSIF ((x0 = TRUE) AND  (x1 = TRUE) AND  (x2 = FALSE) AND  (t0.Q = FALSE)) THEN 
        cstate58 := 2630; y0 := FALSE; y1 := FALSE; t0_start := FALSE; 
    ELSIF ((x0 = TRUE) AND  (x1 = TRUE) AND  (x2 = FALSE) AND  (t0.Q = TRUE)) THEN 
        cstate58 := 2626; y0 := FALSE; y1 := FALSE; t0_start := FALSE; 
    ELSIF ((x0 = TRUE) AND  (x1 = TRUE) AND  (x2 = TRUE) AND  (t0.Q = FALSE)) THEN 
        cstate58 := 2566; y0 := FALSE; y1 := FALSE; t0_start := TRUE; t0_up := FALSE; 
    ELSIF ((x0 = TRUE) AND  (x1 = TRUE) AND  (x2 = TRUE) AND  (t0.Q = TRUE)) THEN 
        cstate58 := 2562; y0 := FALSE; y1 := FALSE; t0_start := TRUE; t0_up := FALSE; 
    END_IF;
6358:
    IF ((x0 = FALSE) AND  (x1 = FALSE) AND  (x2 = FALSE) AND  (t0.Q = FALSE)) THEN 
        cstate58 := 6358; y0 := FALSE; y1 := TRUE; t0_start := FALSE; 
    ELSIF ((x0 = FALSE) AND  (x1 = FALSE) AND  (x2 = FALSE) AND  (t0.Q = TRUE)) THEN 
        cstate58 := 6346; y0 := FALSE; y1 := TRUE; t0_start := FALSE; 
    ELSIF ((x0 = FALSE) AND  (x1 = FALSE) AND  (x2 = TRUE) AND  (t0.Q = FALSE)) THEN 
        cstate58 := 6488; y0 := FALSE; y1 := TRUE; t0_start := TRUE; t0_up := FALSE; 
    ELSIF ((x0 = FALSE) AND  (x1 = FALSE) AND  (x2 = TRUE) AND  (t0.Q = TRUE)) THEN 
        cstate58 := 6476; y0 := FALSE; y1 := TRUE; t0_start := TRUE; t0_up := FALSE; 
    ELSIF ((x0 = FALSE) AND  (x1 = TRUE) AND  (x2 = FALSE) AND  (t0.Q = FALSE)) THEN 
        cstate58 := 6340; y0 := FALSE; y1 := FALSE; t0_start := FALSE; 
    ELSIF ((x0 = FALSE) AND  (x1 = TRUE) AND  (x2 = FALSE) AND  (t0.Q = TRUE)) THEN 
        cstate58 := 6338; y0 := FALSE; y1 := FALSE; t0_start := FALSE; 
    ELSIF ((x0 = FALSE) AND  (x1 = TRUE) AND  (x2 = TRUE) AND  (t0.Q = FALSE)) THEN 
        cstate58 := 6468; y0 := FALSE; y1 := FALSE; t0_start := TRUE; t0_up := FALSE; 
    ELSIF ((x0 = FALSE) AND  (x1 = TRUE) AND  (x2 = TRUE) AND  (t0.Q = TRUE)) THEN 
        cstate58 := 6466; y0 := FALSE; y1 := FALSE; t0_start := TRUE; t0_up := FALSE; 
    ELSIF ((x0 = TRUE) AND  (x1 = FALSE) AND  (x2 = FALSE) AND  (t0.Q = FALSE)) THEN 
        cstate58 := 4168; y0 := TRUE; y1 := FALSE; t0_start := FALSE; 
    ELSIF ((x0 = TRUE) AND  (x1 = FALSE) AND  (x2 = FALSE) AND  (t0.Q = TRUE)) THEN 
        cstate58 := 4162; y0 := TRUE; y1 := FALSE; t0_start := FALSE; 
    ELSIF ((x0 = TRUE) AND  (x1 = FALSE) AND  (x2 = TRUE) AND  (t0.Q = FALSE)) THEN 
        cstate58 := 2760; y0 := FALSE; y1 := FALSE; t0_start := TRUE; t0_up := FALSE; 
    ELSIF ((x0 = TRUE) AND  (x1 = FALSE) AND  (x2 = TRUE) AND  (t0.Q = TRUE)) THEN 
        cstate58 := 2754; y0 := FALSE; y1 := FALSE; t0_start := TRUE; t0_up := FALSE; 
    ELSIF ((x0 = TRUE) AND  (x1 = TRUE) AND  (x2 = FALSE) AND  (t0.Q = FALSE)) THEN 
        cstate58 := 4678; y0 := TRUE; y1 := FALSE; t0_start := FALSE; 
    ELSIF ((x0 = TRUE) AND  (x1 = TRUE) AND  (x2 = FALSE) AND  (t0.Q = TRUE)) THEN 
        cstate58 := 4674; y0 := TRUE; y1 := FALSE; t0_start := FALSE; 
    ELSIF ((x0 = TRUE) AND  (x1 = TRUE) AND  (x2 = TRUE) AND  (t0.Q = FALSE)) THEN 
        cstate58 := 2566; y0 := FALSE; y1 := FALSE; t0_start := TRUE; t0_up := FALSE; 
    ELSIF ((x0 = TRUE) AND  (x1 = TRUE) AND  (x2 = TRUE) AND  (t0.Q = TRUE)) THEN 
        cstate58 := 2562; y0 := FALSE; y1 := FALSE; t0_start := TRUE; t0_up := FALSE; 
    END_IF;
2754:
    IF ((x0 = FALSE) AND  (x1 = FALSE) AND  (x2 = FALSE) AND  (t0.Q = FALSE)) THEN 
        cstate58 := 6404; y0 := FALSE; y1 := FALSE; t0_start := FALSE; 
    ELSIF ((x0 = FALSE) AND  (x1 = FALSE) AND  (x2 = FALSE) AND  (t0.Q = TRUE)) THEN 
        cstate58 := 6338; y0 := FALSE; y1 := FALSE; t0_start := FALSE; 
    ELSIF ((x0 = FALSE) AND  (x1 = FALSE) AND  (x2 = TRUE) AND  (t0.Q = FALSE)) THEN 
        cstate58 := 6468; y0 := FALSE; y1 := FALSE; t0_start := FALSE; 
    ELSIF ((x0 = FALSE) AND  (x1 = FALSE) AND  (x2 = TRUE) AND  (t0.Q = TRUE)) THEN 
        cstate58 := 6530; y0 := FALSE; y1 := FALSE; t0_start := FALSE; 
    ELSIF ((x0 = FALSE) AND  (x1 = TRUE) AND  (x2 = FALSE) AND  (t0.Q = FALSE)) THEN 
        cstate58 := 6404; y0 := FALSE; y1 := FALSE; t0_start := FALSE; 
    ELSIF ((x0 = FALSE) AND  (x1 = TRUE) AND  (x2 = FALSE) AND  (t0.Q = TRUE)) THEN 
        cstate58 := 6338; y0 := FALSE; y1 := FALSE; t0_start := FALSE; 
    ELSIF ((x0 = FALSE) AND  (x1 = TRUE) AND  (x2 = TRUE) AND  (t0.Q = FALSE)) THEN 
        cstate58 := 6468; y0 := FALSE; y1 := FALSE; t0_start := FALSE; 
    ELSIF ((x0 = FALSE) AND  (x1 = TRUE) AND  (x2 = TRUE) AND  (t0.Q = TRUE)) THEN 
        cstate58 := 6530; y0 := FALSE; y1 := FALSE; t0_start := FALSE; 
    ELSIF ((x0 = TRUE) AND  (x1 = FALSE) AND  (x2 = FALSE) AND  (t0.Q = FALSE)) THEN 
        cstate58 := 2184; y0 := FALSE; y1 := FALSE; t0_start := FALSE; 
    ELSIF ((x0 = TRUE) AND  (x1 = FALSE) AND  (x2 = FALSE) AND  (t0.Q = TRUE)) THEN 
        cstate58 := 2114; y0 := FALSE; y1 := FALSE; t0_start := FALSE; 
    ELSIF ((x0 = TRUE) AND  (x1 = FALSE) AND  (x2 = TRUE) AND  (t0.Q = FALSE)) THEN 
        cstate58 := 2760; y0 := FALSE; y1 := FALSE; t0_start := FALSE; 
    ELSIF ((x0 = TRUE) AND  (x1 = FALSE) AND  (x2 = TRUE) AND  (t0.Q = TRUE)) THEN 
        cstate58 := 2818; y0 := FALSE; y1 := FALSE; t0_start := FALSE; 
    ELSIF ((x0 = TRUE) AND  (x1 = TRUE) AND  (x2 = FALSE) AND  (t0.Q = FALSE)) THEN 
        cstate58 := 2694; y0 := FALSE; y1 := FALSE; t0_start := FALSE; 
    ELSIF ((x0 = TRUE) AND  (x1 = TRUE) AND  (x2 = FALSE) AND  (t0.Q = TRUE)) THEN 
        cstate58 := 2626; y0 := FALSE; y1 := FALSE; t0_start := FALSE; 
    ELSIF ((x0 = TRUE) AND  (x1 = TRUE) AND  (x2 = TRUE) AND  (t0.Q = FALSE)) THEN 
        cstate58 := 2566; y0 := FALSE; y1 := FALSE; t0_start := FALSE; 
    ELSIF ((x0 = TRUE) AND  (x1 = TRUE) AND  (x2 = TRUE) AND  (t0.Q = TRUE)) THEN 
        cstate58 := 2498; y0 := FALSE; y1 := FALSE; t0_start := FALSE; 
    END_IF;
6362:
    IF ((x0 = FALSE) AND  (x1 = FALSE) AND  (x2 = FALSE) AND  (t0.Q = FALSE)) THEN 
        cstate58 := 6362; y0 := FALSE; y1 := TRUE; t0_start := FALSE; 
    ELSIF ((x0 = FALSE) AND  (x1 = FALSE) AND  (x2 = FALSE) AND  (t0.Q = TRUE)) THEN 
        cstate58 := 6350; y0 := FALSE; y1 := TRUE; t0_start := FALSE; 
    ELSIF ((x0 = FALSE) AND  (x1 = FALSE) AND  (x2 = TRUE) AND  (t0.Q = FALSE)) THEN 
        cstate58 := 6492; y0 := FALSE; y1 := TRUE; t0_start := TRUE; t0_up := FALSE; 
    ELSIF ((x0 = FALSE) AND  (x1 = FALSE) AND  (x2 = TRUE) AND  (t0.Q = TRUE)) THEN 
        cstate58 := 6480; y0 := FALSE; y1 := TRUE; t0_start := TRUE; t0_up := FALSE; 
    ELSIF ((x0 = FALSE) AND  (x1 = TRUE) AND  (x2 = FALSE) AND  (t0.Q = FALSE)) THEN 
        cstate58 := 6340; y0 := FALSE; y1 := FALSE; t0_start := FALSE; 
    ELSIF ((x0 = FALSE) AND  (x1 = TRUE) AND  (x2 = FALSE) AND  (t0.Q = TRUE)) THEN 
        cstate58 := 6338; y0 := FALSE; y1 := FALSE; t0_start := FALSE; 
    ELSIF ((x0 = FALSE) AND  (x1 = TRUE) AND  (x2 = TRUE) AND  (t0.Q = FALSE)) THEN 
        cstate58 := 6468; y0 := FALSE; y1 := FALSE; t0_start := TRUE; t0_up := FALSE; 
    ELSIF ((x0 = FALSE) AND  (x1 = TRUE) AND  (x2 = TRUE) AND  (t0.Q = TRUE)) THEN 
        cstate58 := 6466; y0 := FALSE; y1 := FALSE; t0_start := TRUE; t0_up := FALSE; 
    ELSIF ((x0 = TRUE) AND  (x1 = FALSE) AND  (x2 = FALSE) AND  (t0.Q = FALSE)) THEN 
        cstate58 := 4168; y0 := TRUE; y1 := FALSE; t0_start := FALSE; 
    ELSIF ((x0 = TRUE) AND  (x1 = FALSE) AND  (x2 = FALSE) AND  (t0.Q = TRUE)) THEN 
        cstate58 := 4162; y0 := TRUE; y1 := FALSE; t0_start := FALSE; 
    ELSIF ((x0 = TRUE) AND  (x1 = FALSE) AND  (x2 = TRUE) AND  (t0.Q = FALSE)) THEN 
        cstate58 := 2760; y0 := FALSE; y1 := FALSE; t0_start := TRUE; t0_up := FALSE; 
    ELSIF ((x0 = TRUE) AND  (x1 = FALSE) AND  (x2 = TRUE) AND  (t0.Q = TRUE)) THEN 
        cstate58 := 2754; y0 := FALSE; y1 := FALSE; t0_start := TRUE; t0_up := FALSE; 
    ELSIF ((x0 = TRUE) AND  (x1 = TRUE) AND  (x2 = FALSE) AND  (t0.Q = FALSE)) THEN 
        cstate58 := 4678; y0 := TRUE; y1 := FALSE; t0_start := FALSE; 
    ELSIF ((x0 = TRUE) AND  (x1 = TRUE) AND  (x2 = FALSE) AND  (t0.Q = TRUE)) THEN 
        cstate58 := 4674; y0 := TRUE; y1 := FALSE; t0_start := FALSE; 
    ELSIF ((x0 = TRUE) AND  (x1 = TRUE) AND  (x2 = TRUE) AND  (t0.Q = FALSE)) THEN 
        cstate58 := 2566; y0 := FALSE; y1 := FALSE; t0_start := TRUE; t0_up := FALSE; 
    ELSIF ((x0 = TRUE) AND  (x1 = TRUE) AND  (x2 = TRUE) AND  (t0.Q = TRUE)) THEN 
        cstate58 := 2562; y0 := FALSE; y1 := FALSE; t0_start := TRUE; t0_up := FALSE; 
    END_IF;
6404:
    IF ((x0 = FALSE) AND  (x1 = FALSE) AND  (x2 = FALSE) AND  (t0.Q = FALSE)) THEN 
        cstate58 := 6404; y0 := FALSE; y1 := FALSE; t0_start := FALSE; 
    ELSIF ((x0 = FALSE) AND  (x1 = FALSE) AND  (x2 = FALSE) AND  (t0.Q = TRUE)) THEN 
        cstate58 := 6346; y0 := FALSE; y1 := TRUE; t0_start := FALSE; 
    ELSIF ((x0 = FALSE) AND  (x1 = FALSE) AND  (x2 = TRUE) AND  (t0.Q = FALSE)) THEN 
        cstate58 := 6468; y0 := FALSE; y1 := FALSE; t0_start := TRUE; t0_up := FALSE; 
    ELSIF ((x0 = FALSE) AND  (x1 = FALSE) AND  (x2 = TRUE) AND  (t0.Q = TRUE)) THEN 
        cstate58 := 6476; y0 := FALSE; y1 := TRUE; t0_start := TRUE; t0_up := FALSE; 
    ELSIF ((x0 = FALSE) AND  (x1 = TRUE) AND  (x2 = FALSE) AND  (t0.Q = FALSE)) THEN 
        cstate58 := 6404; y0 := FALSE; y1 := FALSE; t0_start := FALSE; 
    ELSIF ((x0 = FALSE) AND  (x1 = TRUE) AND  (x2 = FALSE) AND  (t0.Q = TRUE)) THEN 
        cstate58 := 6338; y0 := FALSE; y1 := FALSE; t0_start := FALSE; 
    ELSIF ((x0 = FALSE) AND  (x1 = TRUE) AND  (x2 = TRUE) AND  (t0.Q = FALSE)) THEN 
        cstate58 := 6468; y0 := FALSE; y1 := FALSE; t0_start := TRUE; t0_up := FALSE; 
    ELSIF ((x0 = FALSE) AND  (x1 = TRUE) AND  (x2 = TRUE) AND  (t0.Q = TRUE)) THEN 
        cstate58 := 6466; y0 := FALSE; y1 := FALSE; t0_start := TRUE; t0_up := FALSE; 
    ELSIF ((x0 = TRUE) AND  (x1 = FALSE) AND  (x2 = FALSE) AND  (t0.Q = FALSE)) THEN 
        cstate58 := 4232; y0 := TRUE; y1 := FALSE; t0_start := FALSE; 
    ELSIF ((x0 = TRUE) AND  (x1 = FALSE) AND  (x2 = FALSE) AND  (t0.Q = TRUE)) THEN 
        cstate58 := 4162; y0 := TRUE; y1 := FALSE; t0_start := FALSE; 
    ELSIF ((x0 = TRUE) AND  (x1 = FALSE) AND  (x2 = TRUE) AND  (t0.Q = FALSE)) THEN 
        cstate58 := 2760; y0 := FALSE; y1 := FALSE; t0_start := TRUE; t0_up := FALSE; 
    ELSIF ((x0 = TRUE) AND  (x1 = FALSE) AND  (x2 = TRUE) AND  (t0.Q = TRUE)) THEN 
        cstate58 := 2754; y0 := FALSE; y1 := FALSE; t0_start := TRUE; t0_up := FALSE; 
    ELSIF ((x0 = TRUE) AND  (x1 = TRUE) AND  (x2 = FALSE) AND  (t0.Q = FALSE)) THEN 
        cstate58 := 4742; y0 := TRUE; y1 := FALSE; t0_start := FALSE; 
    ELSIF ((x0 = TRUE) AND  (x1 = TRUE) AND  (x2 = FALSE) AND  (t0.Q = TRUE)) THEN 
        cstate58 := 4674; y0 := TRUE; y1 := FALSE; t0_start := FALSE; 
    ELSIF ((x0 = TRUE) AND  (x1 = TRUE) AND  (x2 = TRUE) AND  (t0.Q = FALSE)) THEN 
        cstate58 := 2566; y0 := FALSE; y1 := FALSE; t0_start := TRUE; t0_up := FALSE; 
    ELSIF ((x0 = TRUE) AND  (x1 = TRUE) AND  (x2 = TRUE) AND  (t0.Q = TRUE)) THEN 
        cstate58 := 2562; y0 := FALSE; y1 := FALSE; t0_start := TRUE; t0_up := FALSE; 
    END_IF;
0:
    IF ((x0 = FALSE) AND  (x1 = FALSE) AND  (x2 = FALSE) AND  (t0.Q = FALSE)) THEN 
        cstate58 := 1220; y0 := FALSE; y1 := FALSE; t0_start := FALSE; 
    ELSIF ((x0 = FALSE) AND  (x1 = FALSE) AND  (x2 = FALSE) AND  (t0.Q = TRUE)) THEN 
        cstate58 := 1218; y0 := FALSE; y1 := FALSE; t0_start := FALSE; 
    ELSIF ((x0 = FALSE) AND  (x1 = FALSE) AND  (x2 = TRUE) AND  (t0.Q = FALSE)) THEN 
        cstate58 := 1412; y0 := FALSE; y1 := FALSE; t0_start := FALSE; 
    ELSIF ((x0 = FALSE) AND  (x1 = FALSE) AND  (x2 = TRUE) AND  (t0.Q = TRUE)) THEN 
        cstate58 := 1410; y0 := FALSE; y1 := FALSE; t0_start := FALSE; 
    ELSIF ((x0 = FALSE) AND  (x1 = TRUE) AND  (x2 = FALSE) AND  (t0.Q = FALSE)) THEN 
        cstate58 := 1220; y0 := FALSE; y1 := FALSE; t0_start := FALSE; 
    ELSIF ((x0 = FALSE) AND  (x1 = TRUE) AND  (x2 = FALSE) AND  (t0.Q = TRUE)) THEN 
        cstate58 := 1218; y0 := FALSE; y1 := FALSE; t0_start := FALSE; 
    ELSIF ((x0 = FALSE) AND  (x1 = TRUE) AND  (x2 = TRUE) AND  (t0.Q = FALSE)) THEN 
        cstate58 := 1412; y0 := FALSE; y1 := FALSE; t0_start := FALSE; 
    ELSIF ((x0 = FALSE) AND  (x1 = TRUE) AND  (x2 = TRUE) AND  (t0.Q = TRUE)) THEN 
        cstate58 := 1410; y0 := FALSE; y1 := FALSE; t0_start := FALSE; 
    ELSIF ((x0 = TRUE) AND  (x1 = FALSE) AND  (x2 = FALSE) AND  (t0.Q = FALSE)) THEN 
        cstate58 := 3144; y0 := FALSE; y1 := FALSE; t0_start := FALSE; 
    ELSIF ((x0 = TRUE) AND  (x1 = FALSE) AND  (x2 = FALSE) AND  (t0.Q = TRUE)) THEN 
        cstate58 := 3138; y0 := FALSE; y1 := FALSE; t0_start := FALSE; 
    ELSIF ((x0 = TRUE) AND  (x1 = FALSE) AND  (x2 = TRUE) AND  (t0.Q = FALSE)) THEN 
        cstate58 := 3848; y0 := FALSE; y1 := FALSE; t0_start := FALSE; 
    ELSIF ((x0 = TRUE) AND  (x1 = FALSE) AND  (x2 = TRUE) AND  (t0.Q = TRUE)) THEN 
        cstate58 := 3842; y0 := FALSE; y1 := FALSE; t0_start := FALSE; 
    ELSIF ((x0 = TRUE) AND  (x1 = TRUE) AND  (x2 = FALSE) AND  (t0.Q = FALSE)) THEN 
        cstate58 := 2630; y0 := FALSE; y1 := FALSE; t0_start := FALSE; 
    ELSIF ((x0 = TRUE) AND  (x1 = TRUE) AND  (x2 = FALSE) AND  (t0.Q = TRUE)) THEN 
        cstate58 := 2626; y0 := FALSE; y1 := FALSE; t0_start := FALSE; 
    ELSIF ((x0 = TRUE) AND  (x1 = TRUE) AND  (x2 = TRUE) AND  (t0.Q = FALSE)) THEN 
        cstate58 := 2502; y0 := FALSE; y1 := FALSE; t0_start := FALSE; 
    ELSIF ((x0 = TRUE) AND  (x1 = TRUE) AND  (x2 = TRUE) AND  (t0.Q = TRUE)) THEN 
        cstate58 := 2498; y0 := FALSE; y1 := FALSE; t0_start := FALSE; 
    END_IF;
6366:
    IF ((x0 = FALSE) AND  (x1 = FALSE) AND  (x2 = FALSE) AND  (t0.Q = FALSE)) THEN 
        cstate58 := 6366; y0 := FALSE; y1 := TRUE; t0_start := FALSE; 
    ELSIF ((x0 = FALSE) AND  (x1 = FALSE) AND  (x2 = FALSE) AND  (t0.Q = TRUE)) THEN 
        cstate58 := 6354; y0 := FALSE; y1 := TRUE; t0_start := FALSE; 
    ELSIF ((x0 = FALSE) AND  (x1 = FALSE) AND  (x2 = TRUE) AND  (t0.Q = FALSE)) THEN 
        cstate58 := 6496; y0 := FALSE; y1 := TRUE; t0_start := TRUE; t0_up := FALSE; 
    ELSIF ((x0 = FALSE) AND  (x1 = FALSE) AND  (x2 = TRUE) AND  (t0.Q = TRUE)) THEN 
        cstate58 := 6484; y0 := FALSE; y1 := TRUE; t0_start := TRUE; t0_up := FALSE; 
    ELSIF ((x0 = FALSE) AND  (x1 = TRUE) AND  (x2 = FALSE) AND  (t0.Q = FALSE)) THEN 
        cstate58 := 6340; y0 := FALSE; y1 := FALSE; t0_start := FALSE; 
    ELSIF ((x0 = FALSE) AND  (x1 = TRUE) AND  (x2 = FALSE) AND  (t0.Q = TRUE)) THEN 
        cstate58 := 6338; y0 := FALSE; y1 := FALSE; t0_start := FALSE; 
    ELSIF ((x0 = FALSE) AND  (x1 = TRUE) AND  (x2 = TRUE) AND  (t0.Q = FALSE)) THEN 
        cstate58 := 6468; y0 := FALSE; y1 := FALSE; t0_start := TRUE; t0_up := FALSE; 
    ELSIF ((x0 = FALSE) AND  (x1 = TRUE) AND  (x2 = TRUE) AND  (t0.Q = TRUE)) THEN 
        cstate58 := 6466; y0 := FALSE; y1 := FALSE; t0_start := TRUE; t0_up := FALSE; 
    ELSIF ((x0 = TRUE) AND  (x1 = FALSE) AND  (x2 = FALSE) AND  (t0.Q = FALSE)) THEN 
        cstate58 := 4168; y0 := TRUE; y1 := FALSE; t0_start := FALSE; 
    ELSIF ((x0 = TRUE) AND  (x1 = FALSE) AND  (x2 = FALSE) AND  (t0.Q = TRUE)) THEN 
        cstate58 := 4162; y0 := TRUE; y1 := FALSE; t0_start := FALSE; 
    ELSIF ((x0 = TRUE) AND  (x1 = FALSE) AND  (x2 = TRUE) AND  (t0.Q = FALSE)) THEN 
        cstate58 := 2760; y0 := FALSE; y1 := FALSE; t0_start := TRUE; t0_up := FALSE; 
    ELSIF ((x0 = TRUE) AND  (x1 = FALSE) AND  (x2 = TRUE) AND  (t0.Q = TRUE)) THEN 
        cstate58 := 2754; y0 := FALSE; y1 := FALSE; t0_start := TRUE; t0_up := FALSE; 
    ELSIF ((x0 = TRUE) AND  (x1 = TRUE) AND  (x2 = FALSE) AND  (t0.Q = FALSE)) THEN 
        cstate58 := 4678; y0 := TRUE; y1 := FALSE; t0_start := FALSE; 
    ELSIF ((x0 = TRUE) AND  (x1 = TRUE) AND  (x2 = FALSE) AND  (t0.Q = TRUE)) THEN 
        cstate58 := 4674; y0 := TRUE; y1 := FALSE; t0_start := FALSE; 
    ELSIF ((x0 = TRUE) AND  (x1 = TRUE) AND  (x2 = TRUE) AND  (t0.Q = FALSE)) THEN 
        cstate58 := 2566; y0 := FALSE; y1 := FALSE; t0_start := TRUE; t0_up := FALSE; 
    ELSIF ((x0 = TRUE) AND  (x1 = TRUE) AND  (x2 = TRUE) AND  (t0.Q = TRUE)) THEN 
        cstate58 := 2562; y0 := FALSE; y1 := FALSE; t0_start := TRUE; t0_up := FALSE; 
    END_IF;
2760:
    IF ((x0 = FALSE) AND  (x1 = FALSE) AND  (x2 = FALSE) AND  (t0.Q = FALSE)) THEN 
        cstate58 := 6404; y0 := FALSE; y1 := FALSE; t0_start := FALSE; 
    ELSIF ((x0 = FALSE) AND  (x1 = FALSE) AND  (x2 = FALSE) AND  (t0.Q = TRUE)) THEN 
        cstate58 := 6354; y0 := FALSE; y1 := TRUE; t0_start := FALSE; 
    ELSIF ((x0 = FALSE) AND  (x1 = FALSE) AND  (x2 = TRUE) AND  (t0.Q = FALSE)) THEN 
        cstate58 := 6468; y0 := FALSE; y1 := FALSE; t0_start := FALSE; 
    ELSIF ((x0 = FALSE) AND  (x1 = FALSE) AND  (x2 = TRUE) AND  (t0.Q = TRUE)) THEN 
        cstate58 := 6546; y0 := FALSE; y1 := TRUE; t0_start := FALSE; 
    ELSIF ((x0 = FALSE) AND  (x1 = TRUE) AND  (x2 = FALSE) AND  (t0.Q = FALSE)) THEN 
        cstate58 := 6404; y0 := FALSE; y1 := FALSE; t0_start := FALSE; 
    ELSIF ((x0 = FALSE) AND  (x1 = TRUE) AND  (x2 = FALSE) AND  (t0.Q = TRUE)) THEN 
        cstate58 := 6338; y0 := FALSE; y1 := FALSE; t0_start := FALSE; 
    ELSIF ((x0 = FALSE) AND  (x1 = TRUE) AND  (x2 = TRUE) AND  (t0.Q = FALSE)) THEN 
        cstate58 := 6468; y0 := FALSE; y1 := FALSE; t0_start := FALSE; 
    ELSIF ((x0 = FALSE) AND  (x1 = TRUE) AND  (x2 = TRUE) AND  (t0.Q = TRUE)) THEN 
        cstate58 := 6530; y0 := FALSE; y1 := FALSE; t0_start := FALSE; 
    ELSIF ((x0 = TRUE) AND  (x1 = FALSE) AND  (x2 = FALSE) AND  (t0.Q = FALSE)) THEN 
        cstate58 := 2184; y0 := FALSE; y1 := FALSE; t0_start := FALSE; 
    ELSIF ((x0 = TRUE) AND  (x1 = FALSE) AND  (x2 = FALSE) AND  (t0.Q = TRUE)) THEN 
        cstate58 := 2114; y0 := FALSE; y1 := FALSE; t0_start := FALSE; 
    ELSIF ((x0 = TRUE) AND  (x1 = FALSE) AND  (x2 = TRUE) AND  (t0.Q = FALSE)) THEN 
        cstate58 := 2760; y0 := FALSE; y1 := FALSE; t0_start := FALSE; 
    ELSIF ((x0 = TRUE) AND  (x1 = FALSE) AND  (x2 = TRUE) AND  (t0.Q = TRUE)) THEN 
        cstate58 := 2818; y0 := FALSE; y1 := FALSE; t0_start := FALSE; 
    ELSIF ((x0 = TRUE) AND  (x1 = TRUE) AND  (x2 = FALSE) AND  (t0.Q = FALSE)) THEN 
        cstate58 := 2694; y0 := FALSE; y1 := FALSE; t0_start := FALSE; 
    ELSIF ((x0 = TRUE) AND  (x1 = TRUE) AND  (x2 = FALSE) AND  (t0.Q = TRUE)) THEN 
        cstate58 := 2626; y0 := FALSE; y1 := FALSE; t0_start := FALSE; 
    ELSIF ((x0 = TRUE) AND  (x1 = TRUE) AND  (x2 = TRUE) AND  (t0.Q = FALSE)) THEN 
        cstate58 := 2566; y0 := FALSE; y1 := FALSE; t0_start := FALSE; 
    ELSIF ((x0 = TRUE) AND  (x1 = TRUE) AND  (x2 = TRUE) AND  (t0.Q = TRUE)) THEN 
        cstate58 := 2498; y0 := FALSE; y1 := FALSE; t0_start := FALSE; 
    END_IF;
6554:
    IF ((x0 = FALSE) AND  (x1 = FALSE) AND  (x2 = FALSE) AND  (t0.Q = FALSE)) THEN 
        cstate58 := 6362; y0 := FALSE; y1 := TRUE; t0_start := FALSE; 
    ELSIF ((x0 = FALSE) AND  (x1 = FALSE) AND  (x2 = FALSE) AND  (t0.Q = TRUE)) THEN 
        cstate58 := 6350; y0 := FALSE; y1 := TRUE; t0_start := FALSE; 
    ELSIF ((x0 = FALSE) AND  (x1 = FALSE) AND  (x2 = TRUE) AND  (t0.Q = FALSE)) THEN 
        cstate58 := 6554; y0 := FALSE; y1 := TRUE; t0_start := FALSE; 
    ELSIF ((x0 = FALSE) AND  (x1 = FALSE) AND  (x2 = TRUE) AND  (t0.Q = TRUE)) THEN 
        cstate58 := 6542; y0 := FALSE; y1 := TRUE; t0_start := FALSE; 
    ELSIF ((x0 = FALSE) AND  (x1 = TRUE) AND  (x2 = FALSE) AND  (t0.Q = FALSE)) THEN 
        cstate58 := 6340; y0 := FALSE; y1 := FALSE; t0_start := FALSE; 
    ELSIF ((x0 = FALSE) AND  (x1 = TRUE) AND  (x2 = FALSE) AND  (t0.Q = TRUE)) THEN 
        cstate58 := 6338; y0 := FALSE; y1 := FALSE; t0_start := FALSE; 
    ELSIF ((x0 = FALSE) AND  (x1 = TRUE) AND  (x2 = TRUE) AND  (t0.Q = FALSE)) THEN 
        cstate58 := 6532; y0 := FALSE; y1 := FALSE; t0_start := FALSE; 
    ELSIF ((x0 = FALSE) AND  (x1 = TRUE) AND  (x2 = TRUE) AND  (t0.Q = TRUE)) THEN 
        cstate58 := 6530; y0 := FALSE; y1 := FALSE; t0_start := FALSE; 
    ELSIF ((x0 = TRUE) AND  (x1 = FALSE) AND  (x2 = FALSE) AND  (t0.Q = FALSE)) THEN 
        cstate58 := 4168; y0 := TRUE; y1 := FALSE; t0_start := FALSE; 
    ELSIF ((x0 = TRUE) AND  (x1 = FALSE) AND  (x2 = FALSE) AND  (t0.Q = TRUE)) THEN 
        cstate58 := 4162; y0 := TRUE; y1 := FALSE; t0_start := FALSE; 
    ELSIF ((x0 = TRUE) AND  (x1 = FALSE) AND  (x2 = TRUE) AND  (t0.Q = FALSE)) THEN 
        cstate58 := 2824; y0 := FALSE; y1 := FALSE; t0_start := FALSE; 
    ELSIF ((x0 = TRUE) AND  (x1 = FALSE) AND  (x2 = TRUE) AND  (t0.Q = TRUE)) THEN 
        cstate58 := 2818; y0 := FALSE; y1 := FALSE; t0_start := FALSE; 
    ELSIF ((x0 = TRUE) AND  (x1 = TRUE) AND  (x2 = FALSE) AND  (t0.Q = FALSE)) THEN 
        cstate58 := 4678; y0 := TRUE; y1 := FALSE; t0_start := FALSE; 
    ELSIF ((x0 = TRUE) AND  (x1 = TRUE) AND  (x2 = FALSE) AND  (t0.Q = TRUE)) THEN 
        cstate58 := 4674; y0 := TRUE; y1 := FALSE; t0_start := FALSE; 
    ELSIF ((x0 = TRUE) AND  (x1 = TRUE) AND  (x2 = TRUE) AND  (t0.Q = FALSE)) THEN 
        cstate58 := 2502; y0 := FALSE; y1 := FALSE; t0_start := FALSE; 
    ELSIF ((x0 = TRUE) AND  (x1 = TRUE) AND  (x2 = TRUE) AND  (t0.Q = TRUE)) THEN 
        cstate58 := 2498; y0 := FALSE; y1 := FALSE; t0_start := FALSE; 
    END_IF;
3144:
    IF ((x0 = FALSE) AND  (x1 = FALSE) AND  (x2 = FALSE) AND  (t0.Q = FALSE)) THEN 
        cstate58 := 7364; y0 := FALSE; y1 := FALSE; t0_start := FALSE; 
    ELSIF ((x0 = FALSE) AND  (x1 = FALSE) AND  (x2 = FALSE) AND  (t0.Q = TRUE)) THEN 
        cstate58 := 7378; y0 := FALSE; y1 := TRUE; t0_start := FALSE; 
    ELSIF ((x0 = FALSE) AND  (x1 = FALSE) AND  (x2 = TRUE) AND  (t0.Q = FALSE)) THEN 
        cstate58 := 7492; y0 := FALSE; y1 := FALSE; t0_start := TRUE; t0_up := FALSE; 
    ELSIF ((x0 = FALSE) AND  (x1 = FALSE) AND  (x2 = TRUE) AND  (t0.Q = TRUE)) THEN 
        cstate58 := 7508; y0 := FALSE; y1 := TRUE; t0_start := TRUE; t0_up := FALSE; 
    ELSIF ((x0 = FALSE) AND  (x1 = TRUE) AND  (x2 = FALSE) AND  (t0.Q = FALSE)) THEN 
        cstate58 := 6340; y0 := FALSE; y1 := FALSE; t0_start := FALSE; 
    ELSIF ((x0 = FALSE) AND  (x1 = TRUE) AND  (x2 = FALSE) AND  (t0.Q = TRUE)) THEN 
        cstate58 := 6338; y0 := FALSE; y1 := FALSE; t0_start := FALSE; 
    ELSIF ((x0 = FALSE) AND  (x1 = TRUE) AND  (x2 = TRUE) AND  (t0.Q = FALSE)) THEN 
        cstate58 := 6468; y0 := FALSE; y1 := FALSE; t0_start := TRUE; t0_up := FALSE; 
    ELSIF ((x0 = FALSE) AND  (x1 = TRUE) AND  (x2 = TRUE) AND  (t0.Q = TRUE)) THEN 
        cstate58 := 6466; y0 := FALSE; y1 := FALSE; t0_start := TRUE; t0_up := FALSE; 
    ELSIF ((x0 = TRUE) AND  (x1 = FALSE) AND  (x2 = FALSE) AND  (t0.Q = FALSE)) THEN 
        cstate58 := 3144; y0 := FALSE; y1 := FALSE; t0_start := FALSE; 
    ELSIF ((x0 = TRUE) AND  (x1 = FALSE) AND  (x2 = FALSE) AND  (t0.Q = TRUE)) THEN 
        cstate58 := 3138; y0 := FALSE; y1 := FALSE; t0_start := FALSE; 
    ELSIF ((x0 = TRUE) AND  (x1 = FALSE) AND  (x2 = TRUE) AND  (t0.Q = FALSE)) THEN 
        cstate58 := 3784; y0 := FALSE; y1 := FALSE; t0_start := TRUE; t0_up := FALSE; 
    ELSIF ((x0 = TRUE) AND  (x1 = FALSE) AND  (x2 = TRUE) AND  (t0.Q = TRUE)) THEN 
        cstate58 := 3778; y0 := FALSE; y1 := FALSE; t0_start := TRUE; t0_up := FALSE; 
    ELSIF ((x0 = TRUE) AND  (x1 = TRUE) AND  (x2 = FALSE) AND  (t0.Q = FALSE)) THEN 
        cstate58 := 2630; y0 := FALSE; y1 := FALSE; t0_start := FALSE; 
    ELSIF ((x0 = TRUE) AND  (x1 = TRUE) AND  (x2 = FALSE) AND  (t0.Q = TRUE)) THEN 
        cstate58 := 2626; y0 := FALSE; y1 := FALSE; t0_start := FALSE; 
    ELSIF ((x0 = TRUE) AND  (x1 = TRUE) AND  (x2 = TRUE) AND  (t0.Q = FALSE)) THEN 
        cstate58 := 2566; y0 := FALSE; y1 := FALSE; t0_start := TRUE; t0_up := FALSE; 
    ELSIF ((x0 = TRUE) AND  (x1 = TRUE) AND  (x2 = TRUE) AND  (t0.Q = TRUE)) THEN 
        cstate58 := 2562; y0 := FALSE; y1 := FALSE; t0_start := TRUE; t0_up := FALSE; 
    END_IF;
7556:
    IF ((x0 = FALSE) AND  (x1 = FALSE) AND  (x2 = FALSE) AND  (t0.Q = FALSE)) THEN 
        cstate58 := 7364; y0 := FALSE; y1 := FALSE; t0_start := FALSE; 
    ELSIF ((x0 = FALSE) AND  (x1 = FALSE) AND  (x2 = FALSE) AND  (t0.Q = TRUE)) THEN 
        cstate58 := 7370; y0 := FALSE; y1 := TRUE; t0_start := FALSE; 
    ELSIF ((x0 = FALSE) AND  (x1 = FALSE) AND  (x2 = TRUE) AND  (t0.Q = FALSE)) THEN 
        cstate58 := 7556; y0 := FALSE; y1 := FALSE; t0_start := FALSE; 
    ELSIF ((x0 = FALSE) AND  (x1 = FALSE) AND  (x2 = TRUE) AND  (t0.Q = TRUE)) THEN 
        cstate58 := 7562; y0 := FALSE; y1 := TRUE; t0_start := FALSE; 
    ELSIF ((x0 = FALSE) AND  (x1 = TRUE) AND  (x2 = FALSE) AND  (t0.Q = FALSE)) THEN 
        cstate58 := 6340; y0 := FALSE; y1 := FALSE; t0_start := FALSE; 
    ELSIF ((x0 = FALSE) AND  (x1 = TRUE) AND  (x2 = FALSE) AND  (t0.Q = TRUE)) THEN 
        cstate58 := 6338; y0 := FALSE; y1 := FALSE; t0_start := FALSE; 
    ELSIF ((x0 = FALSE) AND  (x1 = TRUE) AND  (x2 = TRUE) AND  (t0.Q = FALSE)) THEN 
        cstate58 := 6532; y0 := FALSE; y1 := FALSE; t0_start := FALSE; 
    ELSIF ((x0 = FALSE) AND  (x1 = TRUE) AND  (x2 = TRUE) AND  (t0.Q = TRUE)) THEN 
        cstate58 := 6530; y0 := FALSE; y1 := FALSE; t0_start := FALSE; 
    ELSIF ((x0 = TRUE) AND  (x1 = FALSE) AND  (x2 = FALSE) AND  (t0.Q = FALSE)) THEN 
        cstate58 := 5192; y0 := TRUE; y1 := FALSE; t0_start := FALSE; 
    ELSIF ((x0 = TRUE) AND  (x1 = FALSE) AND  (x2 = FALSE) AND  (t0.Q = TRUE)) THEN 
        cstate58 := 5186; y0 := TRUE; y1 := FALSE; t0_start := FALSE; 
    ELSIF ((x0 = TRUE) AND  (x1 = FALSE) AND  (x2 = TRUE) AND  (t0.Q = FALSE)) THEN 
        cstate58 := 3848; y0 := FALSE; y1 := FALSE; t0_start := FALSE; 
    ELSIF ((x0 = TRUE) AND  (x1 = FALSE) AND  (x2 = TRUE) AND  (t0.Q = TRUE)) THEN 
        cstate58 := 3842; y0 := FALSE; y1 := FALSE; t0_start := FALSE; 
    ELSIF ((x0 = TRUE) AND  (x1 = TRUE) AND  (x2 = FALSE) AND  (t0.Q = FALSE)) THEN 
        cstate58 := 4678; y0 := TRUE; y1 := FALSE; t0_start := FALSE; 
    ELSIF ((x0 = TRUE) AND  (x1 = TRUE) AND  (x2 = FALSE) AND  (t0.Q = TRUE)) THEN 
        cstate58 := 4674; y0 := TRUE; y1 := FALSE; t0_start := FALSE; 
    ELSIF ((x0 = TRUE) AND  (x1 = TRUE) AND  (x2 = TRUE) AND  (t0.Q = FALSE)) THEN 
        cstate58 := 2502; y0 := FALSE; y1 := FALSE; t0_start := FALSE; 
    ELSIF ((x0 = TRUE) AND  (x1 = TRUE) AND  (x2 = TRUE) AND  (t0.Q = TRUE)) THEN 
        cstate58 := 2498; y0 := FALSE; y1 := FALSE; t0_start := FALSE; 
    END_IF;
7554:
    IF ((x0 = FALSE) AND  (x1 = FALSE) AND  (x2 = FALSE) AND  (t0.Q = FALSE)) THEN 
        cstate58 := 7364; y0 := FALSE; y1 := FALSE; t0_start := FALSE; 
    ELSIF ((x0 = FALSE) AND  (x1 = FALSE) AND  (x2 = FALSE) AND  (t0.Q = TRUE)) THEN 
        cstate58 := 7362; y0 := FALSE; y1 := FALSE; t0_start := FALSE; 
    ELSIF ((x0 = FALSE) AND  (x1 = FALSE) AND  (x2 = TRUE) AND  (t0.Q = FALSE)) THEN 
        cstate58 := 7556; y0 := FALSE; y1 := FALSE; t0_start := FALSE; 
    ELSIF ((x0 = FALSE) AND  (x1 = FALSE) AND  (x2 = TRUE) AND  (t0.Q = TRUE)) THEN 
        cstate58 := 7554; y0 := FALSE; y1 := FALSE; t0_start := FALSE; 
    ELSIF ((x0 = FALSE) AND  (x1 = TRUE) AND  (x2 = FALSE) AND  (t0.Q = FALSE)) THEN 
        cstate58 := 6340; y0 := FALSE; y1 := FALSE; t0_start := FALSE; 
    ELSIF ((x0 = FALSE) AND  (x1 = TRUE) AND  (x2 = FALSE) AND  (t0.Q = TRUE)) THEN 
        cstate58 := 6338; y0 := FALSE; y1 := FALSE; t0_start := FALSE; 
    ELSIF ((x0 = FALSE) AND  (x1 = TRUE) AND  (x2 = TRUE) AND  (t0.Q = FALSE)) THEN 
        cstate58 := 6532; y0 := FALSE; y1 := FALSE; t0_start := FALSE; 
    ELSIF ((x0 = FALSE) AND  (x1 = TRUE) AND  (x2 = TRUE) AND  (t0.Q = TRUE)) THEN 
        cstate58 := 6530; y0 := FALSE; y1 := FALSE; t0_start := FALSE; 
    ELSIF ((x0 = TRUE) AND  (x1 = FALSE) AND  (x2 = FALSE) AND  (t0.Q = FALSE)) THEN 
        cstate58 := 5192; y0 := TRUE; y1 := FALSE; t0_start := FALSE; 
    ELSIF ((x0 = TRUE) AND  (x1 = FALSE) AND  (x2 = FALSE) AND  (t0.Q = TRUE)) THEN 
        cstate58 := 5186; y0 := TRUE; y1 := FALSE; t0_start := FALSE; 
    ELSIF ((x0 = TRUE) AND  (x1 = FALSE) AND  (x2 = TRUE) AND  (t0.Q = FALSE)) THEN 
        cstate58 := 3848; y0 := FALSE; y1 := FALSE; t0_start := FALSE; 
    ELSIF ((x0 = TRUE) AND  (x1 = FALSE) AND  (x2 = TRUE) AND  (t0.Q = TRUE)) THEN 
        cstate58 := 3842; y0 := FALSE; y1 := FALSE; t0_start := FALSE; 
    ELSIF ((x0 = TRUE) AND  (x1 = TRUE) AND  (x2 = FALSE) AND  (t0.Q = FALSE)) THEN 
        cstate58 := 4678; y0 := TRUE; y1 := FALSE; t0_start := FALSE; 
    ELSIF ((x0 = TRUE) AND  (x1 = TRUE) AND  (x2 = FALSE) AND  (t0.Q = TRUE)) THEN 
        cstate58 := 4674; y0 := TRUE; y1 := FALSE; t0_start := FALSE; 
    ELSIF ((x0 = TRUE) AND  (x1 = TRUE) AND  (x2 = TRUE) AND  (t0.Q = FALSE)) THEN 
        cstate58 := 2502; y0 := FALSE; y1 := FALSE; t0_start := FALSE; 
    ELSIF ((x0 = TRUE) AND  (x1 = TRUE) AND  (x2 = TRUE) AND  (t0.Q = TRUE)) THEN 
        cstate58 := 2498; y0 := FALSE; y1 := FALSE; t0_start := FALSE; 
    END_IF;
6550:
    IF ((x0 = FALSE) AND  (x1 = FALSE) AND  (x2 = FALSE) AND  (t0.Q = FALSE)) THEN 
        cstate58 := 6358; y0 := FALSE; y1 := TRUE; t0_start := FALSE; 
    ELSIF ((x0 = FALSE) AND  (x1 = FALSE) AND  (x2 = FALSE) AND  (t0.Q = TRUE)) THEN 
        cstate58 := 6346; y0 := FALSE; y1 := TRUE; t0_start := FALSE; 
    ELSIF ((x0 = FALSE) AND  (x1 = FALSE) AND  (x2 = TRUE) AND  (t0.Q = FALSE)) THEN 
        cstate58 := 6550; y0 := FALSE; y1 := TRUE; t0_start := FALSE; 
    ELSIF ((x0 = FALSE) AND  (x1 = FALSE) AND  (x2 = TRUE) AND  (t0.Q = TRUE)) THEN 
        cstate58 := 6538; y0 := FALSE; y1 := TRUE; t0_start := FALSE; 
    ELSIF ((x0 = FALSE) AND  (x1 = TRUE) AND  (x2 = FALSE) AND  (t0.Q = FALSE)) THEN 
        cstate58 := 6340; y0 := FALSE; y1 := FALSE; t0_start := FALSE; 
    ELSIF ((x0 = FALSE) AND  (x1 = TRUE) AND  (x2 = FALSE) AND  (t0.Q = TRUE)) THEN 
        cstate58 := 6338; y0 := FALSE; y1 := FALSE; t0_start := FALSE; 
    ELSIF ((x0 = FALSE) AND  (x1 = TRUE) AND  (x2 = TRUE) AND  (t0.Q = FALSE)) THEN 
        cstate58 := 6532; y0 := FALSE; y1 := FALSE; t0_start := FALSE; 
    ELSIF ((x0 = FALSE) AND  (x1 = TRUE) AND  (x2 = TRUE) AND  (t0.Q = TRUE)) THEN 
        cstate58 := 6530; y0 := FALSE; y1 := FALSE; t0_start := FALSE; 
    ELSIF ((x0 = TRUE) AND  (x1 = FALSE) AND  (x2 = FALSE) AND  (t0.Q = FALSE)) THEN 
        cstate58 := 4168; y0 := TRUE; y1 := FALSE; t0_start := FALSE; 
    ELSIF ((x0 = TRUE) AND  (x1 = FALSE) AND  (x2 = FALSE) AND  (t0.Q = TRUE)) THEN 
        cstate58 := 4162; y0 := TRUE; y1 := FALSE; t0_start := FALSE; 
    ELSIF ((x0 = TRUE) AND  (x1 = FALSE) AND  (x2 = TRUE) AND  (t0.Q = FALSE)) THEN 
        cstate58 := 2824; y0 := FALSE; y1 := FALSE; t0_start := FALSE; 
    ELSIF ((x0 = TRUE) AND  (x1 = FALSE) AND  (x2 = TRUE) AND  (t0.Q = TRUE)) THEN 
        cstate58 := 2818; y0 := FALSE; y1 := FALSE; t0_start := FALSE; 
    ELSIF ((x0 = TRUE) AND  (x1 = TRUE) AND  (x2 = FALSE) AND  (t0.Q = FALSE)) THEN 
        cstate58 := 4678; y0 := TRUE; y1 := FALSE; t0_start := FALSE; 
    ELSIF ((x0 = TRUE) AND  (x1 = TRUE) AND  (x2 = FALSE) AND  (t0.Q = TRUE)) THEN 
        cstate58 := 4674; y0 := TRUE; y1 := FALSE; t0_start := FALSE; 
    ELSIF ((x0 = TRUE) AND  (x1 = TRUE) AND  (x2 = TRUE) AND  (t0.Q = FALSE)) THEN 
        cstate58 := 2502; y0 := FALSE; y1 := FALSE; t0_start := FALSE; 
    ELSIF ((x0 = TRUE) AND  (x1 = TRUE) AND  (x2 = TRUE) AND  (t0.Q = TRUE)) THEN 
        cstate58 := 2498; y0 := FALSE; y1 := FALSE; t0_start := FALSE; 
    END_IF;
6468:
    IF ((x0 = FALSE) AND  (x1 = FALSE) AND  (x2 = FALSE) AND  (t0.Q = FALSE)) THEN 
        cstate58 := 6404; y0 := FALSE; y1 := FALSE; t0_start := FALSE; 
    ELSIF ((x0 = FALSE) AND  (x1 = FALSE) AND  (x2 = FALSE) AND  (t0.Q = TRUE)) THEN 
        cstate58 := 6346; y0 := FALSE; y1 := TRUE; t0_start := FALSE; 
    ELSIF ((x0 = FALSE) AND  (x1 = FALSE) AND  (x2 = TRUE) AND  (t0.Q = FALSE)) THEN 
        cstate58 := 6468; y0 := FALSE; y1 := FALSE; t0_start := FALSE; 
    ELSIF ((x0 = FALSE) AND  (x1 = FALSE) AND  (x2 = TRUE) AND  (t0.Q = TRUE)) THEN 
        cstate58 := 6538; y0 := FALSE; y1 := TRUE; t0_start := FALSE; 
    ELSIF ((x0 = FALSE) AND  (x1 = TRUE) AND  (x2 = FALSE) AND  (t0.Q = FALSE)) THEN 
        cstate58 := 6404; y0 := FALSE; y1 := FALSE; t0_start := FALSE; 
    ELSIF ((x0 = FALSE) AND  (x1 = TRUE) AND  (x2 = FALSE) AND  (t0.Q = TRUE)) THEN 
        cstate58 := 6338; y0 := FALSE; y1 := FALSE; t0_start := FALSE; 
    ELSIF ((x0 = FALSE) AND  (x1 = TRUE) AND  (x2 = TRUE) AND  (t0.Q = FALSE)) THEN 
        cstate58 := 6468; y0 := FALSE; y1 := FALSE; t0_start := FALSE; 
    ELSIF ((x0 = FALSE) AND  (x1 = TRUE) AND  (x2 = TRUE) AND  (t0.Q = TRUE)) THEN 
        cstate58 := 6530; y0 := FALSE; y1 := FALSE; t0_start := FALSE; 
    ELSIF ((x0 = TRUE) AND  (x1 = FALSE) AND  (x2 = FALSE) AND  (t0.Q = FALSE)) THEN 
        cstate58 := 4232; y0 := TRUE; y1 := FALSE; t0_start := FALSE; 
    ELSIF ((x0 = TRUE) AND  (x1 = FALSE) AND  (x2 = FALSE) AND  (t0.Q = TRUE)) THEN 
        cstate58 := 4162; y0 := TRUE; y1 := FALSE; t0_start := FALSE; 
    ELSIF ((x0 = TRUE) AND  (x1 = FALSE) AND  (x2 = TRUE) AND  (t0.Q = FALSE)) THEN 
        cstate58 := 2760; y0 := FALSE; y1 := FALSE; t0_start := FALSE; 
    ELSIF ((x0 = TRUE) AND  (x1 = FALSE) AND  (x2 = TRUE) AND  (t0.Q = TRUE)) THEN 
        cstate58 := 2818; y0 := FALSE; y1 := FALSE; t0_start := FALSE; 
    ELSIF ((x0 = TRUE) AND  (x1 = TRUE) AND  (x2 = FALSE) AND  (t0.Q = FALSE)) THEN 
        cstate58 := 4742; y0 := TRUE; y1 := FALSE; t0_start := FALSE; 
    ELSIF ((x0 = TRUE) AND  (x1 = TRUE) AND  (x2 = FALSE) AND  (t0.Q = TRUE)) THEN 
        cstate58 := 4674; y0 := TRUE; y1 := FALSE; t0_start := FALSE; 
    ELSIF ((x0 = TRUE) AND  (x1 = TRUE) AND  (x2 = TRUE) AND  (t0.Q = FALSE)) THEN 
        cstate58 := 2566; y0 := FALSE; y1 := FALSE; t0_start := FALSE; 
    ELSIF ((x0 = TRUE) AND  (x1 = TRUE) AND  (x2 = TRUE) AND  (t0.Q = TRUE)) THEN 
        cstate58 := 2498; y0 := FALSE; y1 := FALSE; t0_start := FALSE; 
    END_IF;
5256:
    IF ((x0 = FALSE) AND  (x1 = FALSE) AND  (x2 = FALSE) AND  (t0.Q = FALSE)) THEN 
        cstate58 := 9476; y0 := TRUE; y1 := FALSE; t0_start := FALSE; 
    ELSIF ((x0 = FALSE) AND  (x1 = FALSE) AND  (x2 = FALSE) AND  (t0.Q = TRUE)) THEN 
        cstate58 := 9410; y0 := TRUE; y1 := FALSE; t0_start := FALSE; 
    ELSIF ((x0 = FALSE) AND  (x1 = FALSE) AND  (x2 = TRUE) AND  (t0.Q = FALSE)) THEN 
        cstate58 := 7492; y0 := FALSE; y1 := FALSE; t0_start := TRUE; t0_up := FALSE; 
    ELSIF ((x0 = FALSE) AND  (x1 = FALSE) AND  (x2 = TRUE) AND  (t0.Q = TRUE)) THEN 
        cstate58 := 7508; y0 := FALSE; y1 := TRUE; t0_start := TRUE; t0_up := FALSE; 
    ELSIF ((x0 = FALSE) AND  (x1 = TRUE) AND  (x2 = FALSE) AND  (t0.Q = FALSE)) THEN 
        cstate58 := 8452; y0 := TRUE; y1 := FALSE; t0_start := FALSE; 
    ELSIF ((x0 = FALSE) AND  (x1 = TRUE) AND  (x2 = FALSE) AND  (t0.Q = TRUE)) THEN 
        cstate58 := 8386; y0 := TRUE; y1 := FALSE; t0_start := FALSE; 
    ELSIF ((x0 = FALSE) AND  (x1 = TRUE) AND  (x2 = TRUE) AND  (t0.Q = FALSE)) THEN 
        cstate58 := 6468; y0 := FALSE; y1 := FALSE; t0_start := TRUE; t0_up := FALSE; 
    ELSIF ((x0 = FALSE) AND  (x1 = TRUE) AND  (x2 = TRUE) AND  (t0.Q = TRUE)) THEN 
        cstate58 := 6466; y0 := FALSE; y1 := FALSE; t0_start := TRUE; t0_up := FALSE; 
    ELSIF ((x0 = TRUE) AND  (x1 = FALSE) AND  (x2 = FALSE) AND  (t0.Q = FALSE)) THEN 
        cstate58 := 5256; y0 := TRUE; y1 := FALSE; t0_start := FALSE; 
    ELSIF ((x0 = TRUE) AND  (x1 = FALSE) AND  (x2 = FALSE) AND  (t0.Q = TRUE)) THEN 
        cstate58 := 5186; y0 := TRUE; y1 := FALSE; t0_start := FALSE; 
    ELSIF ((x0 = TRUE) AND  (x1 = FALSE) AND  (x2 = TRUE) AND  (t0.Q = FALSE)) THEN 
        cstate58 := 3784; y0 := FALSE; y1 := FALSE; t0_start := TRUE; t0_up := FALSE; 
    ELSIF ((x0 = TRUE) AND  (x1 = FALSE) AND  (x2 = TRUE) AND  (t0.Q = TRUE)) THEN 
        cstate58 := 3778; y0 := FALSE; y1 := FALSE; t0_start := TRUE; t0_up := FALSE; 
    ELSIF ((x0 = TRUE) AND  (x1 = TRUE) AND  (x2 = FALSE) AND  (t0.Q = FALSE)) THEN 
        cstate58 := 4742; y0 := TRUE; y1 := FALSE; t0_start := FALSE; 
    ELSIF ((x0 = TRUE) AND  (x1 = TRUE) AND  (x2 = FALSE) AND  (t0.Q = TRUE)) THEN 
        cstate58 := 4674; y0 := TRUE; y1 := FALSE; t0_start := FALSE; 
    ELSIF ((x0 = TRUE) AND  (x1 = TRUE) AND  (x2 = TRUE) AND  (t0.Q = FALSE)) THEN 
        cstate58 := 2566; y0 := FALSE; y1 := FALSE; t0_start := TRUE; t0_up := FALSE; 
    ELSIF ((x0 = TRUE) AND  (x1 = TRUE) AND  (x2 = TRUE) AND  (t0.Q = TRUE)) THEN 
        cstate58 := 2562; y0 := FALSE; y1 := FALSE; t0_start := TRUE; t0_up := FALSE; 
    END_IF;
8388:
    IF ((x0 = FALSE) AND  ( TRUE ) AND  (x2 = FALSE) AND  (t0.Q = FALSE)) THEN 
        cstate58 := 8388; y0 := TRUE; y1 := FALSE; t0_start := FALSE; 
    ELSIF ((x0 = FALSE) AND  ( TRUE ) AND  (x2 = FALSE) AND  (t0.Q = TRUE)) THEN 
        cstate58 := 8386; y0 := TRUE; y1 := FALSE; t0_start := FALSE; 
    ELSIF ((x0 = FALSE) AND  (x1 = FALSE) AND  (x2 = TRUE) AND  (t0.Q = FALSE)) THEN 
        cstate58 := 6468; y0 := FALSE; y1 := FALSE; t0_start := TRUE; t0_up := FALSE; 
    ELSIF ((x0 = FALSE) AND  (x1 = FALSE) AND  (x2 = TRUE) AND  (t0.Q = TRUE)) THEN 
        cstate58 := 6476; y0 := FALSE; y1 := TRUE; t0_start := TRUE; t0_up := FALSE; 
    ELSIF ((x0 = FALSE) AND  (x1 = TRUE) AND  (x2 = TRUE) AND  (t0.Q = FALSE)) THEN 
        cstate58 := 6468; y0 := FALSE; y1 := FALSE; t0_start := TRUE; t0_up := FALSE; 
    ELSIF ((x0 = FALSE) AND  (x1 = TRUE) AND  (x2 = TRUE) AND  (t0.Q = TRUE)) THEN 
        cstate58 := 6466; y0 := FALSE; y1 := FALSE; t0_start := TRUE; t0_up := FALSE; 
    ELSIF ((x0 = TRUE) AND  (x1 = FALSE) AND  (x2 = FALSE) AND  (t0.Q = FALSE)) THEN 
        cstate58 := 4168; y0 := TRUE; y1 := FALSE; t0_start := FALSE; 
    ELSIF ((x0 = TRUE) AND  (x1 = FALSE) AND  (x2 = FALSE) AND  (t0.Q = TRUE)) THEN 
        cstate58 := 4162; y0 := TRUE; y1 := FALSE; t0_start := FALSE; 
    ELSIF ((x0 = TRUE) AND  (x1 = FALSE) AND  (x2 = TRUE) AND  (t0.Q = FALSE)) THEN 
        cstate58 := 2760; y0 := FALSE; y1 := FALSE; t0_start := TRUE; t0_up := FALSE; 
    ELSIF ((x0 = TRUE) AND  (x1 = FALSE) AND  (x2 = TRUE) AND  (t0.Q = TRUE)) THEN 
        cstate58 := 2754; y0 := FALSE; y1 := FALSE; t0_start := TRUE; t0_up := FALSE; 
    ELSIF ((x0 = TRUE) AND  (x1 = TRUE) AND  (x2 = FALSE) AND  (t0.Q = FALSE)) THEN 
        cstate58 := 4678; y0 := TRUE; y1 := FALSE; t0_start := FALSE; 
    ELSIF ((x0 = TRUE) AND  (x1 = TRUE) AND  (x2 = FALSE) AND  (t0.Q = TRUE)) THEN 
        cstate58 := 4674; y0 := TRUE; y1 := FALSE; t0_start := FALSE; 
    ELSIF ((x0 = TRUE) AND  (x1 = TRUE) AND  (x2 = TRUE) AND  (t0.Q = FALSE)) THEN 
        cstate58 := 2566; y0 := FALSE; y1 := FALSE; t0_start := TRUE; t0_up := FALSE; 
    ELSIF ((x0 = TRUE) AND  (x1 = TRUE) AND  (x2 = TRUE) AND  (t0.Q = TRUE)) THEN 
        cstate58 := 2562; y0 := FALSE; y1 := FALSE; t0_start := TRUE; t0_up := FALSE; 
    END_IF;
3848:
    IF ((x0 = FALSE) AND  (x1 = FALSE) AND  (x2 = FALSE) AND  (t0.Q = FALSE)) THEN 
        cstate58 := 7364; y0 := FALSE; y1 := FALSE; t0_start := FALSE; 
    ELSIF ((x0 = FALSE) AND  (x1 = FALSE) AND  (x2 = FALSE) AND  (t0.Q = TRUE)) THEN 
        cstate58 := 7378; y0 := FALSE; y1 := TRUE; t0_start := FALSE; 
    ELSIF ((x0 = FALSE) AND  (x1 = FALSE) AND  (x2 = TRUE) AND  (t0.Q = FALSE)) THEN 
        cstate58 := 7556; y0 := FALSE; y1 := FALSE; t0_start := FALSE; 
    ELSIF ((x0 = FALSE) AND  (x1 = FALSE) AND  (x2 = TRUE) AND  (t0.Q = TRUE)) THEN 
        cstate58 := 7570; y0 := FALSE; y1 := TRUE; t0_start := FALSE; 
    ELSIF ((x0 = FALSE) AND  (x1 = TRUE) AND  (x2 = FALSE) AND  (t0.Q = FALSE)) THEN 
        cstate58 := 6340; y0 := FALSE; y1 := FALSE; t0_start := FALSE; 
    ELSIF ((x0 = FALSE) AND  (x1 = TRUE) AND  (x2 = FALSE) AND  (t0.Q = TRUE)) THEN 
        cstate58 := 6338; y0 := FALSE; y1 := FALSE; t0_start := FALSE; 
    ELSIF ((x0 = FALSE) AND  (x1 = TRUE) AND  (x2 = TRUE) AND  (t0.Q = FALSE)) THEN 
        cstate58 := 6532; y0 := FALSE; y1 := FALSE; t0_start := FALSE; 
    ELSIF ((x0 = FALSE) AND  (x1 = TRUE) AND  (x2 = TRUE) AND  (t0.Q = TRUE)) THEN 
        cstate58 := 6530; y0 := FALSE; y1 := FALSE; t0_start := FALSE; 
    ELSIF ((x0 = TRUE) AND  (x1 = FALSE) AND  (x2 = FALSE) AND  (t0.Q = FALSE)) THEN 
        cstate58 := 3144; y0 := FALSE; y1 := FALSE; t0_start := FALSE; 
    ELSIF ((x0 = TRUE) AND  (x1 = FALSE) AND  (x2 = FALSE) AND  (t0.Q = TRUE)) THEN 
        cstate58 := 3138; y0 := FALSE; y1 := FALSE; t0_start := FALSE; 
    ELSIF ((x0 = TRUE) AND  (x1 = FALSE) AND  (x2 = TRUE) AND  (t0.Q = FALSE)) THEN 
        cstate58 := 3848; y0 := FALSE; y1 := FALSE; t0_start := FALSE; 
    ELSIF ((x0 = TRUE) AND  (x1 = FALSE) AND  (x2 = TRUE) AND  (t0.Q = TRUE)) THEN 
        cstate58 := 3842; y0 := FALSE; y1 := FALSE; t0_start := FALSE; 
    ELSIF ((x0 = TRUE) AND  (x1 = TRUE) AND  (x2 = FALSE) AND  (t0.Q = FALSE)) THEN 
        cstate58 := 2630; y0 := FALSE; y1 := FALSE; t0_start := FALSE; 
    ELSIF ((x0 = TRUE) AND  (x1 = TRUE) AND  (x2 = FALSE) AND  (t0.Q = TRUE)) THEN 
        cstate58 := 2626; y0 := FALSE; y1 := FALSE; t0_start := FALSE; 
    ELSIF ((x0 = TRUE) AND  (x1 = TRUE) AND  (x2 = TRUE) AND  (t0.Q = FALSE)) THEN 
        cstate58 := 2502; y0 := FALSE; y1 := FALSE; t0_start := FALSE; 
    ELSIF ((x0 = TRUE) AND  (x1 = TRUE) AND  (x2 = TRUE) AND  (t0.Q = TRUE)) THEN 
        cstate58 := 2498; y0 := FALSE; y1 := FALSE; t0_start := FALSE; 
    END_IF;
1430:
    IF ((x0 = FALSE) AND  (x1 = FALSE) AND  (x2 = FALSE) AND  (t0.Q = FALSE)) THEN 
        cstate58 := 1238; y0 := FALSE; y1 := TRUE; t0_start := FALSE; 
    ELSIF ((x0 = FALSE) AND  (x1 = FALSE) AND  (x2 = FALSE) AND  (t0.Q = TRUE)) THEN 
        cstate58 := 1226; y0 := FALSE; y1 := TRUE; t0_start := FALSE; 
    ELSIF ((x0 = FALSE) AND  (x1 = FALSE) AND  (x2 = TRUE) AND  (t0.Q = FALSE)) THEN 
        cstate58 := 1430; y0 := FALSE; y1 := TRUE; t0_start := FALSE; 
    ELSIF ((x0 = FALSE) AND  (x1 = FALSE) AND  (x2 = TRUE) AND  (t0.Q = TRUE)) THEN 
        cstate58 := 1418; y0 := FALSE; y1 := TRUE; t0_start := FALSE; 
    ELSIF ((x0 = FALSE) AND  (x1 = TRUE) AND  (x2 = FALSE) AND  (t0.Q = FALSE)) THEN 
        cstate58 := 1220; y0 := FALSE; y1 := FALSE; t0_start := FALSE; 
    ELSIF ((x0 = FALSE) AND  (x1 = TRUE) AND  (x2 = FALSE) AND  (t0.Q = TRUE)) THEN 
        cstate58 := 1218; y0 := FALSE; y1 := FALSE; t0_start := FALSE; 
    ELSIF ((x0 = FALSE) AND  (x1 = TRUE) AND  (x2 = TRUE) AND  (t0.Q = FALSE)) THEN 
        cstate58 := 1412; y0 := FALSE; y1 := FALSE; t0_start := FALSE; 
    ELSIF ((x0 = FALSE) AND  (x1 = TRUE) AND  (x2 = TRUE) AND  (t0.Q = TRUE)) THEN 
        cstate58 := 1410; y0 := FALSE; y1 := FALSE; t0_start := FALSE; 
    ELSIF ((x0 = TRUE) AND  (x1 = FALSE) AND  (x2 = FALSE) AND  (t0.Q = FALSE)) THEN 
        cstate58 := 5192; y0 := TRUE; y1 := FALSE; t0_start := FALSE; 
    ELSIF ((x0 = TRUE) AND  (x1 = FALSE) AND  (x2 = FALSE) AND  (t0.Q = TRUE)) THEN 
        cstate58 := 5186; y0 := TRUE; y1 := FALSE; t0_start := FALSE; 
    ELSIF ((x0 = TRUE) AND  (x1 = FALSE) AND  (x2 = TRUE) AND  (t0.Q = FALSE)) THEN 
        cstate58 := 3848; y0 := FALSE; y1 := FALSE; t0_start := FALSE; 
    ELSIF ((x0 = TRUE) AND  (x1 = FALSE) AND  (x2 = TRUE) AND  (t0.Q = TRUE)) THEN 
        cstate58 := 3842; y0 := FALSE; y1 := FALSE; t0_start := FALSE; 
    ELSIF ((x0 = TRUE) AND  (x1 = TRUE) AND  (x2 = FALSE) AND  (t0.Q = FALSE)) THEN 
        cstate58 := 4678; y0 := TRUE; y1 := FALSE; t0_start := FALSE; 
    ELSIF ((x0 = TRUE) AND  (x1 = TRUE) AND  (x2 = FALSE) AND  (t0.Q = TRUE)) THEN 
        cstate58 := 4674; y0 := TRUE; y1 := FALSE; t0_start := FALSE; 
    ELSIF ((x0 = TRUE) AND  (x1 = TRUE) AND  (x2 = TRUE) AND  (t0.Q = FALSE)) THEN 
        cstate58 := 2502; y0 := FALSE; y1 := FALSE; t0_start := FALSE; 
    ELSIF ((x0 = TRUE) AND  (x1 = TRUE) AND  (x2 = TRUE) AND  (t0.Q = TRUE)) THEN 
        cstate58 := 2498; y0 := FALSE; y1 := FALSE; t0_start := FALSE; 
    END_IF;
8386:
    IF ((x0 = FALSE) AND  ( TRUE ) AND  (x2 = FALSE) AND  (t0.Q = FALSE)) THEN 
        cstate58 := 8388; y0 := TRUE; y1 := FALSE; t0_start := FALSE; 
    ELSIF ((x0 = FALSE) AND  ( TRUE ) AND  (x2 = FALSE) AND  (t0.Q = TRUE)) THEN 
        cstate58 := 8386; y0 := TRUE; y1 := FALSE; t0_start := FALSE; 
    ELSIF ((x0 = FALSE) AND  (x1 = FALSE) AND  (x2 = TRUE) AND  (t0.Q = FALSE)) THEN 
        cstate58 := 6468; y0 := FALSE; y1 := FALSE; t0_start := TRUE; t0_up := FALSE; 
    ELSIF ((x0 = FALSE) AND  (x1 = FALSE) AND  (x2 = TRUE) AND  (t0.Q = TRUE)) THEN 
        cstate58 := 6466; y0 := FALSE; y1 := FALSE; t0_start := TRUE; t0_up := FALSE; 
    ELSIF ((x0 = FALSE) AND  (x1 = TRUE) AND  (x2 = TRUE) AND  (t0.Q = FALSE)) THEN 
        cstate58 := 6468; y0 := FALSE; y1 := FALSE; t0_start := TRUE; t0_up := FALSE; 
    ELSIF ((x0 = FALSE) AND  (x1 = TRUE) AND  (x2 = TRUE) AND  (t0.Q = TRUE)) THEN 
        cstate58 := 6466; y0 := FALSE; y1 := FALSE; t0_start := TRUE; t0_up := FALSE; 
    ELSIF ((x0 = TRUE) AND  (x1 = FALSE) AND  (x2 = FALSE) AND  (t0.Q = FALSE)) THEN 
        cstate58 := 4168; y0 := TRUE; y1 := FALSE; t0_start := FALSE; 
    ELSIF ((x0 = TRUE) AND  (x1 = FALSE) AND  (x2 = FALSE) AND  (t0.Q = TRUE)) THEN 
        cstate58 := 4162; y0 := TRUE; y1 := FALSE; t0_start := FALSE; 
    ELSIF ((x0 = TRUE) AND  (x1 = FALSE) AND  (x2 = TRUE) AND  (t0.Q = FALSE)) THEN 
        cstate58 := 2760; y0 := FALSE; y1 := FALSE; t0_start := TRUE; t0_up := FALSE; 
    ELSIF ((x0 = TRUE) AND  (x1 = FALSE) AND  (x2 = TRUE) AND  (t0.Q = TRUE)) THEN 
        cstate58 := 2754; y0 := FALSE; y1 := FALSE; t0_start := TRUE; t0_up := FALSE; 
    ELSIF ((x0 = TRUE) AND  (x1 = TRUE) AND  (x2 = FALSE) AND  (t0.Q = FALSE)) THEN 
        cstate58 := 4678; y0 := TRUE; y1 := FALSE; t0_start := FALSE; 
    ELSIF ((x0 = TRUE) AND  (x1 = TRUE) AND  (x2 = FALSE) AND  (t0.Q = TRUE)) THEN 
        cstate58 := 4674; y0 := TRUE; y1 := FALSE; t0_start := FALSE; 
    ELSIF ((x0 = TRUE) AND  (x1 = TRUE) AND  (x2 = TRUE) AND  (t0.Q = FALSE)) THEN 
        cstate58 := 2566; y0 := FALSE; y1 := FALSE; t0_start := TRUE; t0_up := FALSE; 
    ELSIF ((x0 = TRUE) AND  (x1 = TRUE) AND  (x2 = TRUE) AND  (t0.Q = TRUE)) THEN 
        cstate58 := 2562; y0 := FALSE; y1 := FALSE; t0_start := TRUE; t0_up := FALSE; 
    END_IF;
2626:
    IF ((x0 = FALSE) AND  (x1 = FALSE) AND  (x2 = FALSE) AND  (t0.Q = FALSE)) THEN 
        cstate58 := 6340; y0 := FALSE; y1 := FALSE; t0_start := FALSE; 
    ELSIF ((x0 = FALSE) AND  (x1 = FALSE) AND  (x2 = FALSE) AND  (t0.Q = TRUE)) THEN 
        cstate58 := 6338; y0 := FALSE; y1 := FALSE; t0_start := FALSE; 
    ELSIF ((x0 = FALSE) AND  (x1 = FALSE) AND  (x2 = TRUE) AND  (t0.Q = FALSE)) THEN 
        cstate58 := 6468; y0 := FALSE; y1 := FALSE; t0_start := TRUE; t0_up := FALSE; 
    ELSIF ((x0 = FALSE) AND  (x1 = FALSE) AND  (x2 = TRUE) AND  (t0.Q = TRUE)) THEN 
        cstate58 := 6466; y0 := FALSE; y1 := FALSE; t0_start := TRUE; t0_up := FALSE; 
    ELSIF ((x0 = FALSE) AND  (x1 = TRUE) AND  (x2 = FALSE) AND  (t0.Q = FALSE)) THEN 
        cstate58 := 6340; y0 := FALSE; y1 := FALSE; t0_start := FALSE; 
    ELSIF ((x0 = FALSE) AND  (x1 = TRUE) AND  (x2 = FALSE) AND  (t0.Q = TRUE)) THEN 
        cstate58 := 6338; y0 := FALSE; y1 := FALSE; t0_start := FALSE; 
    ELSIF ((x0 = FALSE) AND  (x1 = TRUE) AND  (x2 = TRUE) AND  (t0.Q = FALSE)) THEN 
        cstate58 := 6468; y0 := FALSE; y1 := FALSE; t0_start := TRUE; t0_up := FALSE; 
    ELSIF ((x0 = FALSE) AND  (x1 = TRUE) AND  (x2 = TRUE) AND  (t0.Q = TRUE)) THEN 
        cstate58 := 6466; y0 := FALSE; y1 := FALSE; t0_start := TRUE; t0_up := FALSE; 
    ELSIF ((x0 = TRUE) AND  (x1 = FALSE) AND  (x2 = FALSE) AND  (t0.Q = FALSE)) THEN 
        cstate58 := 2120; y0 := FALSE; y1 := FALSE; t0_start := FALSE; 
    ELSIF ((x0 = TRUE) AND  (x1 = FALSE) AND  (x2 = FALSE) AND  (t0.Q = TRUE)) THEN 
        cstate58 := 2114; y0 := FALSE; y1 := FALSE; t0_start := FALSE; 
    ELSIF ((x0 = TRUE) AND  (x1 = FALSE) AND  (x2 = TRUE) AND  (t0.Q = FALSE)) THEN 
        cstate58 := 2760; y0 := FALSE; y1 := FALSE; t0_start := TRUE; t0_up := FALSE; 
    ELSIF ((x0 = TRUE) AND  (x1 = FALSE) AND  (x2 = TRUE) AND  (t0.Q = TRUE)) THEN 
        cstate58 := 2754; y0 := FALSE; y1 := FALSE; t0_start := TRUE; t0_up := FALSE; 
    ELSIF ((x0 = TRUE) AND  (x1 = TRUE) AND  (x2 = FALSE) AND  (t0.Q = FALSE)) THEN 
        cstate58 := 2630; y0 := FALSE; y1 := FALSE; t0_start := FALSE; 
    ELSIF ((x0 = TRUE) AND  (x1 = TRUE) AND  (x2 = FALSE) AND  (t0.Q = TRUE)) THEN 
        cstate58 := 2626; y0 := FALSE; y1 := FALSE; t0_start := FALSE; 
    ELSIF ((x0 = TRUE) AND  (x1 = TRUE) AND  (x2 = TRUE) AND  (t0.Q = FALSE)) THEN 
        cstate58 := 2566; y0 := FALSE; y1 := FALSE; t0_start := TRUE; t0_up := FALSE; 
    ELSIF ((x0 = TRUE) AND  (x1 = TRUE) AND  (x2 = TRUE) AND  (t0.Q = TRUE)) THEN 
        cstate58 := 2562; y0 := FALSE; y1 := FALSE; t0_start := TRUE; t0_up := FALSE; 
    END_IF;
3842:
    IF ((x0 = FALSE) AND  (x1 = FALSE) AND  (x2 = FALSE) AND  (t0.Q = FALSE)) THEN 
        cstate58 := 7364; y0 := FALSE; y1 := FALSE; t0_start := FALSE; 
    ELSIF ((x0 = FALSE) AND  (x1 = FALSE) AND  (x2 = FALSE) AND  (t0.Q = TRUE)) THEN 
        cstate58 := 7362; y0 := FALSE; y1 := FALSE; t0_start := FALSE; 
    ELSIF ((x0 = FALSE) AND  (x1 = FALSE) AND  (x2 = TRUE) AND  (t0.Q = FALSE)) THEN 
        cstate58 := 7556; y0 := FALSE; y1 := FALSE; t0_start := FALSE; 
    ELSIF ((x0 = FALSE) AND  (x1 = FALSE) AND  (x2 = TRUE) AND  (t0.Q = TRUE)) THEN 
        cstate58 := 7554; y0 := FALSE; y1 := FALSE; t0_start := FALSE; 
    ELSIF ((x0 = FALSE) AND  (x1 = TRUE) AND  (x2 = FALSE) AND  (t0.Q = FALSE)) THEN 
        cstate58 := 6340; y0 := FALSE; y1 := FALSE; t0_start := FALSE; 
    ELSIF ((x0 = FALSE) AND  (x1 = TRUE) AND  (x2 = FALSE) AND  (t0.Q = TRUE)) THEN 
        cstate58 := 6338; y0 := FALSE; y1 := FALSE; t0_start := FALSE; 
    ELSIF ((x0 = FALSE) AND  (x1 = TRUE) AND  (x2 = TRUE) AND  (t0.Q = FALSE)) THEN 
        cstate58 := 6532; y0 := FALSE; y1 := FALSE; t0_start := FALSE; 
    ELSIF ((x0 = FALSE) AND  (x1 = TRUE) AND  (x2 = TRUE) AND  (t0.Q = TRUE)) THEN 
        cstate58 := 6530; y0 := FALSE; y1 := FALSE; t0_start := FALSE; 
    ELSIF ((x0 = TRUE) AND  (x1 = FALSE) AND  (x2 = FALSE) AND  (t0.Q = FALSE)) THEN 
        cstate58 := 3144; y0 := FALSE; y1 := FALSE; t0_start := FALSE; 
    ELSIF ((x0 = TRUE) AND  (x1 = FALSE) AND  (x2 = FALSE) AND  (t0.Q = TRUE)) THEN 
        cstate58 := 3138; y0 := FALSE; y1 := FALSE; t0_start := FALSE; 
    ELSIF ((x0 = TRUE) AND  (x1 = FALSE) AND  (x2 = TRUE) AND  (t0.Q = FALSE)) THEN 
        cstate58 := 3848; y0 := FALSE; y1 := FALSE; t0_start := FALSE; 
    ELSIF ((x0 = TRUE) AND  (x1 = FALSE) AND  (x2 = TRUE) AND  (t0.Q = TRUE)) THEN 
        cstate58 := 3842; y0 := FALSE; y1 := FALSE; t0_start := FALSE; 
    ELSIF ((x0 = TRUE) AND  (x1 = TRUE) AND  (x2 = FALSE) AND  (t0.Q = FALSE)) THEN 
        cstate58 := 2630; y0 := FALSE; y1 := FALSE; t0_start := FALSE; 
    ELSIF ((x0 = TRUE) AND  (x1 = TRUE) AND  (x2 = FALSE) AND  (t0.Q = TRUE)) THEN 
        cstate58 := 2626; y0 := FALSE; y1 := FALSE; t0_start := FALSE; 
    ELSIF ((x0 = TRUE) AND  (x1 = TRUE) AND  (x2 = TRUE) AND  (t0.Q = FALSE)) THEN 
        cstate58 := 2502; y0 := FALSE; y1 := FALSE; t0_start := FALSE; 
    ELSIF ((x0 = TRUE) AND  (x1 = TRUE) AND  (x2 = TRUE) AND  (t0.Q = TRUE)) THEN 
        cstate58 := 2498; y0 := FALSE; y1 := FALSE; t0_start := FALSE; 
    END_IF;
7520:
    IF ((x0 = FALSE) AND  (x1 = FALSE) AND  (x2 = FALSE) AND  (t0.Q = FALSE)) THEN 
        cstate58 := 7456; y0 := FALSE; y1 := TRUE; t0_start := FALSE; 
    ELSIF ((x0 = FALSE) AND  (x1 = FALSE) AND  (x2 = FALSE) AND  (t0.Q = TRUE)) THEN 
        cstate58 := 7378; y0 := FALSE; y1 := TRUE; t0_start := FALSE; 
    ELSIF ((x0 = FALSE) AND  (x1 = FALSE) AND  (x2 = TRUE) AND  (t0.Q = FALSE)) THEN 
        cstate58 := 7520; y0 := FALSE; y1 := TRUE; t0_start := FALSE; 
    ELSIF ((x0 = FALSE) AND  (x1 = FALSE) AND  (x2 = TRUE) AND  (t0.Q = TRUE)) THEN 
        cstate58 := 7570; y0 := FALSE; y1 := TRUE; t0_start := FALSE; 
    ELSIF ((x0 = FALSE) AND  (x1 = TRUE) AND  (x2 = FALSE) AND  (t0.Q = FALSE)) THEN 
        cstate58 := 6404; y0 := FALSE; y1 := FALSE; t0_start := FALSE; 
    ELSIF ((x0 = FALSE) AND  (x1 = TRUE) AND  (x2 = FALSE) AND  (t0.Q = TRUE)) THEN 
        cstate58 := 6338; y0 := FALSE; y1 := FALSE; t0_start := FALSE; 
    ELSIF ((x0 = FALSE) AND  (x1 = TRUE) AND  (x2 = TRUE) AND  (t0.Q = FALSE)) THEN 
        cstate58 := 6468; y0 := FALSE; y1 := FALSE; t0_start := FALSE; 
    ELSIF ((x0 = FALSE) AND  (x1 = TRUE) AND  (x2 = TRUE) AND  (t0.Q = TRUE)) THEN 
        cstate58 := 6530; y0 := FALSE; y1 := FALSE; t0_start := FALSE; 
    ELSIF ((x0 = TRUE) AND  (x1 = FALSE) AND  (x2 = FALSE) AND  (t0.Q = FALSE)) THEN 
        cstate58 := 5256; y0 := TRUE; y1 := FALSE; t0_start := FALSE; 
    ELSIF ((x0 = TRUE) AND  (x1 = FALSE) AND  (x2 = FALSE) AND  (t0.Q = TRUE)) THEN 
        cstate58 := 5186; y0 := TRUE; y1 := FALSE; t0_start := FALSE; 
    ELSIF ((x0 = TRUE) AND  (x1 = FALSE) AND  (x2 = TRUE) AND  (t0.Q = FALSE)) THEN 
        cstate58 := 3784; y0 := FALSE; y1 := FALSE; t0_start := FALSE; 
    ELSIF ((x0 = TRUE) AND  (x1 = FALSE) AND  (x2 = TRUE) AND  (t0.Q = TRUE)) THEN 
        cstate58 := 3842; y0 := FALSE; y1 := FALSE; t0_start := FALSE; 
    ELSIF ((x0 = TRUE) AND  (x1 = TRUE) AND  (x2 = FALSE) AND  (t0.Q = FALSE)) THEN 
        cstate58 := 4742; y0 := TRUE; y1 := FALSE; t0_start := FALSE; 
    ELSIF ((x0 = TRUE) AND  (x1 = TRUE) AND  (x2 = FALSE) AND  (t0.Q = TRUE)) THEN 
        cstate58 := 4674; y0 := TRUE; y1 := FALSE; t0_start := FALSE; 
    ELSIF ((x0 = TRUE) AND  (x1 = TRUE) AND  (x2 = TRUE) AND  (t0.Q = FALSE)) THEN 
        cstate58 := 2566; y0 := FALSE; y1 := FALSE; t0_start := FALSE; 
    ELSIF ((x0 = TRUE) AND  (x1 = TRUE) AND  (x2 = TRUE) AND  (t0.Q = TRUE)) THEN 
        cstate58 := 2498; y0 := FALSE; y1 := FALSE; t0_start := FALSE; 
    END_IF;
6476:
    IF ((x0 = FALSE) AND  (x1 = FALSE) AND  (x2 = FALSE) AND  (t0.Q = FALSE)) THEN 
        cstate58 := 6424; y0 := FALSE; y1 := TRUE; t0_start := FALSE; 
    ELSIF ((x0 = FALSE) AND  (x1 = FALSE) AND  (x2 = FALSE) AND  (t0.Q = TRUE)) THEN 
        cstate58 := 6346; y0 := FALSE; y1 := TRUE; t0_start := FALSE; 
    ELSIF ((x0 = FALSE) AND  (x1 = FALSE) AND  (x2 = TRUE) AND  (t0.Q = FALSE)) THEN 
        cstate58 := 6488; y0 := FALSE; y1 := TRUE; t0_start := FALSE; 
    ELSIF ((x0 = FALSE) AND  (x1 = FALSE) AND  (x2 = TRUE) AND  (t0.Q = TRUE)) THEN 
        cstate58 := 6538; y0 := FALSE; y1 := TRUE; t0_start := FALSE; 
    ELSIF ((x0 = FALSE) AND  (x1 = TRUE) AND  (x2 = FALSE) AND  (t0.Q = FALSE)) THEN 
        cstate58 := 6404; y0 := FALSE; y1 := FALSE; t0_start := FALSE; 
    ELSIF ((x0 = FALSE) AND  (x1 = TRUE) AND  (x2 = FALSE) AND  (t0.Q = TRUE)) THEN 
        cstate58 := 6338; y0 := FALSE; y1 := FALSE; t0_start := FALSE; 
    ELSIF ((x0 = FALSE) AND  (x1 = TRUE) AND  (x2 = TRUE) AND  (t0.Q = FALSE)) THEN 
        cstate58 := 6468; y0 := FALSE; y1 := FALSE; t0_start := FALSE; 
    ELSIF ((x0 = FALSE) AND  (x1 = TRUE) AND  (x2 = TRUE) AND  (t0.Q = TRUE)) THEN 
        cstate58 := 6530; y0 := FALSE; y1 := FALSE; t0_start := FALSE; 
    ELSIF ((x0 = TRUE) AND  (x1 = FALSE) AND  (x2 = FALSE) AND  (t0.Q = FALSE)) THEN 
        cstate58 := 4232; y0 := TRUE; y1 := FALSE; t0_start := FALSE; 
    ELSIF ((x0 = TRUE) AND  (x1 = FALSE) AND  (x2 = FALSE) AND  (t0.Q = TRUE)) THEN 
        cstate58 := 4162; y0 := TRUE; y1 := FALSE; t0_start := FALSE; 
    ELSIF ((x0 = TRUE) AND  (x1 = FALSE) AND  (x2 = TRUE) AND  (t0.Q = FALSE)) THEN 
        cstate58 := 2760; y0 := FALSE; y1 := FALSE; t0_start := FALSE; 
    ELSIF ((x0 = TRUE) AND  (x1 = FALSE) AND  (x2 = TRUE) AND  (t0.Q = TRUE)) THEN 
        cstate58 := 2818; y0 := FALSE; y1 := FALSE; t0_start := FALSE; 
    ELSIF ((x0 = TRUE) AND  (x1 = TRUE) AND  (x2 = FALSE) AND  (t0.Q = FALSE)) THEN 
        cstate58 := 4742; y0 := TRUE; y1 := FALSE; t0_start := FALSE; 
    ELSIF ((x0 = TRUE) AND  (x1 = TRUE) AND  (x2 = FALSE) AND  (t0.Q = TRUE)) THEN 
        cstate58 := 4674; y0 := TRUE; y1 := FALSE; t0_start := FALSE; 
    ELSIF ((x0 = TRUE) AND  (x1 = TRUE) AND  (x2 = TRUE) AND  (t0.Q = FALSE)) THEN 
        cstate58 := 2566; y0 := FALSE; y1 := FALSE; t0_start := FALSE; 
    ELSIF ((x0 = TRUE) AND  (x1 = TRUE) AND  (x2 = TRUE) AND  (t0.Q = TRUE)) THEN 
        cstate58 := 2498; y0 := FALSE; y1 := FALSE; t0_start := FALSE; 
    END_IF;
4232:
    IF ((x0 = FALSE) AND  ( TRUE ) AND  (x2 = FALSE) AND  (t0.Q = FALSE)) THEN 
        cstate58 := 8452; y0 := TRUE; y1 := FALSE; t0_start := FALSE; 
    ELSIF ((x0 = FALSE) AND  ( TRUE ) AND  (x2 = FALSE) AND  (t0.Q = TRUE)) THEN 
        cstate58 := 8386; y0 := TRUE; y1 := FALSE; t0_start := FALSE; 
    ELSIF ((x0 = FALSE) AND  (x1 = FALSE) AND  (x2 = TRUE) AND  (t0.Q = FALSE)) THEN 
        cstate58 := 6468; y0 := FALSE; y1 := FALSE; t0_start := TRUE; t0_up := FALSE; 
    ELSIF ((x0 = FALSE) AND  (x1 = FALSE) AND  (x2 = TRUE) AND  (t0.Q = TRUE)) THEN 
        cstate58 := 6484; y0 := FALSE; y1 := TRUE; t0_start := TRUE; t0_up := FALSE; 
    ELSIF ((x0 = FALSE) AND  (x1 = TRUE) AND  (x2 = TRUE) AND  (t0.Q = FALSE)) THEN 
        cstate58 := 6468; y0 := FALSE; y1 := FALSE; t0_start := TRUE; t0_up := FALSE; 
    ELSIF ((x0 = FALSE) AND  (x1 = TRUE) AND  (x2 = TRUE) AND  (t0.Q = TRUE)) THEN 
        cstate58 := 6466; y0 := FALSE; y1 := FALSE; t0_start := TRUE; t0_up := FALSE; 
    ELSIF ((x0 = TRUE) AND  (x1 = FALSE) AND  (x2 = FALSE) AND  (t0.Q = FALSE)) THEN 
        cstate58 := 4232; y0 := TRUE; y1 := FALSE; t0_start := FALSE; 
    ELSIF ((x0 = TRUE) AND  (x1 = FALSE) AND  (x2 = FALSE) AND  (t0.Q = TRUE)) THEN 
        cstate58 := 4162; y0 := TRUE; y1 := FALSE; t0_start := FALSE; 
    ELSIF ((x0 = TRUE) AND  (x1 = FALSE) AND  (x2 = TRUE) AND  (t0.Q = FALSE)) THEN 
        cstate58 := 2760; y0 := FALSE; y1 := FALSE; t0_start := TRUE; t0_up := FALSE; 
    ELSIF ((x0 = TRUE) AND  (x1 = FALSE) AND  (x2 = TRUE) AND  (t0.Q = TRUE)) THEN 
        cstate58 := 2754; y0 := FALSE; y1 := FALSE; t0_start := TRUE; t0_up := FALSE; 
    ELSIF ((x0 = TRUE) AND  (x1 = TRUE) AND  (x2 = FALSE) AND  (t0.Q = FALSE)) THEN 
        cstate58 := 4742; y0 := TRUE; y1 := FALSE; t0_start := FALSE; 
    ELSIF ((x0 = TRUE) AND  (x1 = TRUE) AND  (x2 = FALSE) AND  (t0.Q = TRUE)) THEN 
        cstate58 := 4674; y0 := TRUE; y1 := FALSE; t0_start := FALSE; 
    ELSIF ((x0 = TRUE) AND  (x1 = TRUE) AND  (x2 = TRUE) AND  (t0.Q = FALSE)) THEN 
        cstate58 := 2566; y0 := FALSE; y1 := FALSE; t0_start := TRUE; t0_up := FALSE; 
    ELSIF ((x0 = TRUE) AND  (x1 = TRUE) AND  (x2 = TRUE) AND  (t0.Q = TRUE)) THEN 
        cstate58 := 2562; y0 := FALSE; y1 := FALSE; t0_start := TRUE; t0_up := FALSE; 
    END_IF;
2630:
    IF ((x0 = FALSE) AND  (x1 = FALSE) AND  (x2 = FALSE) AND  (t0.Q = FALSE)) THEN 
        cstate58 := 6340; y0 := FALSE; y1 := FALSE; t0_start := FALSE; 
    ELSIF ((x0 = FALSE) AND  (x1 = FALSE) AND  (x2 = FALSE) AND  (t0.Q = TRUE)) THEN 
        cstate58 := 6350; y0 := FALSE; y1 := TRUE; t0_start := FALSE; 
    ELSIF ((x0 = FALSE) AND  (x1 = FALSE) AND  (x2 = TRUE) AND  (t0.Q = FALSE)) THEN 
        cstate58 := 6468; y0 := FALSE; y1 := FALSE; t0_start := TRUE; t0_up := FALSE; 
    ELSIF ((x0 = FALSE) AND  (x1 = FALSE) AND  (x2 = TRUE) AND  (t0.Q = TRUE)) THEN 
        cstate58 := 6480; y0 := FALSE; y1 := TRUE; t0_start := TRUE; t0_up := FALSE; 
    ELSIF ((x0 = FALSE) AND  (x1 = TRUE) AND  (x2 = FALSE) AND  (t0.Q = FALSE)) THEN 
        cstate58 := 6340; y0 := FALSE; y1 := FALSE; t0_start := FALSE; 
    ELSIF ((x0 = FALSE) AND  (x1 = TRUE) AND  (x2 = FALSE) AND  (t0.Q = TRUE)) THEN 
        cstate58 := 6338; y0 := FALSE; y1 := FALSE; t0_start := FALSE; 
    ELSIF ((x0 = FALSE) AND  (x1 = TRUE) AND  (x2 = TRUE) AND  (t0.Q = FALSE)) THEN 
        cstate58 := 6468; y0 := FALSE; y1 := FALSE; t0_start := TRUE; t0_up := FALSE; 
    ELSIF ((x0 = FALSE) AND  (x1 = TRUE) AND  (x2 = TRUE) AND  (t0.Q = TRUE)) THEN 
        cstate58 := 6466; y0 := FALSE; y1 := FALSE; t0_start := TRUE; t0_up := FALSE; 
    ELSIF ((x0 = TRUE) AND  (x1 = FALSE) AND  (x2 = FALSE) AND  (t0.Q = FALSE)) THEN 
        cstate58 := 2120; y0 := FALSE; y1 := FALSE; t0_start := FALSE; 
    ELSIF ((x0 = TRUE) AND  (x1 = FALSE) AND  (x2 = FALSE) AND  (t0.Q = TRUE)) THEN 
        cstate58 := 2114; y0 := FALSE; y1 := FALSE; t0_start := FALSE; 
    ELSIF ((x0 = TRUE) AND  (x1 = FALSE) AND  (x2 = TRUE) AND  (t0.Q = FALSE)) THEN 
        cstate58 := 2760; y0 := FALSE; y1 := FALSE; t0_start := TRUE; t0_up := FALSE; 
    ELSIF ((x0 = TRUE) AND  (x1 = FALSE) AND  (x2 = TRUE) AND  (t0.Q = TRUE)) THEN 
        cstate58 := 2754; y0 := FALSE; y1 := FALSE; t0_start := TRUE; t0_up := FALSE; 
